(* PLC project EFBSH-649_PLC, ЗАО "Борисовский завод Металлист" CODESYS CODESYS V3.5 *)
(* stored: creationDateTime 2026-09-25T08:47:37, modificationDateTime 2026-09-25T08:47:37 *)

(* 8 регистров, адрес = 1100 + (индекс-1)*8 *)
TYPE ST_BunkerHmi :
STRUCT
    wSts      : WORD;   (* +0 маски GVL_Const.BS_* *)
    wAlm      : WORD;   (* +1 GVL_Const.BA_SF *)
    wBypass   : WORD;   (* +2 GVL_Const.BY_DVU *)
    uTDvu     : UINT;   (* +3 с *)
    uTRestart : UINT;   (* +4 с *)
    uRes5     : UINT;
    uRes6     : UINT;
    uRes7     : UINT;
END_STRUCT
END_TYPE

TYPE ST_BunkerIn :
STRUCT
    xDVU : BOOL;   (* 1 = верхний уровень *)
    xDNU : BOOL;   (* 1 = продукт на нижнем уровне (для бункера поз.27 - второй датчик) *)
    xSF  : BOOL;   (* станции TORBA: 1 = автомат пульта управления включен *)
END_STRUCT
END_TYPE

TYPE ST_BunkerPar :
STRUCT
    wBypass   : WORD;   (* GVL_Const.BY_DVU - ДВУ отключен *)
    uTDvu     : UINT;   (* задержка срабатывания ДВУ, с *)
    uTRestart : UINT;   (* задержка повторного пуска после снятия ДВУ, с *)
END_STRUCT
END_TYPE

(* Общий блок, %MW0..%MW31 *)
TYPE ST_GlobHmi :
STRUCT
    wCmd        : WORD;  (* +0  маски GVL_Const.G_* *)
    wSts        : WORD;  (* +1  маски GVL_Const.GS_* *)
    wAlm        : WORD;  (* +2  аварийные стопы 1..10 (биты 0..9), 10 пожар, 11 фазы *)
    wWarn       : WORD;  (* +3  маски GVL_Const.GW_* *)
    uHeartbeat  : UINT;  (* +4  счётчик секунд, контроль связи *)
    uTPreStart  : UINT;  (* +5  предпусковой сигнал, с *)
    uTDksGrace  : UINT;  (* +6  разгон до контроля ДКС, с *)
    uTDksPulse  : UINT;  (* +7  нет импульсов ДКС, 0.1 с *)
    uTFcFb      : UINT;  (* +8  нет сигнала работы ПЧ, с *)
    uTFsStart   : UINT;  (* +9  нет статуса фотосепаратора после пуска, с *)
    uTGateMove  : UINT;  (* +10 контроль хода заслонки поз.1, с *)
    uSirenOn    : UINT;  (* +11 1 = аварийная сирена разрешена *)
    uRes        : ARRAY[12..31] OF UINT;
END_STRUCT
END_TYPE

TYPE ST_GlobPar :
STRUCT
    uTPreStart : UINT;
    uTDksGrace : UINT;
    uTDksPulse : UINT;   (* 0.1 с *)
    uTFcFb     : UINT;
    uTFsStart  : UINT;
    uTGateMove : UINT;
    uSirenOn   : UINT;
END_STRUCT
END_TYPE

(* Связь "механизм подаёт на ..." для блокировок и последовательностей *)
TYPE ST_Link :
STRUCT
    iFrom    : INT;    (* индекс механизма-источника *)
    eTo      : INT;    (* GVL_Const.LT_MECH / LT_BUNKER / LT_INVALID *)
    iTo      : INT;    (* индекс механизма или бункера *)
    xProduct : BOOL;   (* TRUE - поток продукта (пауза по ДВУ распространяется назад),
                          FALSE - вспомогательная связь (аспирация, отходы) *)
END_STRUCT
END_TYPE

(* Постоянная конфигурация механизма *)
TYPE ST_MechCfg :
STRUCT
    eKind     : INT;     (* GVL_Const.K_DOL / K_FC / K_GATE / K_FS *)
    xHasQF    : BOOL;    (* контроль автомата защиты (QF/SF) *)
    eDks      : INT;     (* GVL_Const.DKS_NONE / DKS_PULSE / DKS_LEVEL *)
    xHasDSL   : BOOL;    (* датчики сбегания ленты 1 и 2 *)
    xHasDP    : BOOL;    (* датчик подпора *)
    xHasLocal : BOOL;    (* пост местного управления: ключ Авт/Ручн, Пуск, Стоп *)
    xHasEStop : BOOL;    (* аварийный/концевой стоп у механизма *)
    uDefTOn   : UINT;    (* задержка пуска по умолчанию, с *)
    uDefTOff  : UINT;    (* задержка останова по умолчанию, с *)
END_STRUCT
END_TYPE

(* Обмен с панелью по механизму: 16 регистров %MW (только 16-битные поля).
   Адрес = 200 + (индекс-1)*16 + смещение. *)
TYPE ST_MechHmi :
STRUCT
    wCmd           : WORD;  (* +0  команды панели, маски GVL_Const.C_* *)
    wSts           : WORD;  (* +1  состояние, маски GVL_Const.S_* *)
    wAlm           : WORD;  (* +2  аварии (с фиксацией), маски GVL_Const.A_* *)
    wBypass        : WORD;  (* +3  отключение датчиков (запись с паролем) *)
    uTOn           : UINT;  (* +4  задержка пуска, с *)
    uTOff          : UINT;  (* +5  задержка останова, с *)
    uToInterval    : UINT;  (* +6  интервал ТО, ч *)
    uHoursSinceTO  : UINT;  (* +7  наработка после ТО, ч *)
    uHoursTotal    : UINT;  (* +8  наработка всего, ч *)
    uMinutes       : UINT;  (* +9  минуты наработки (0..59) *)
    iState         : INT;   (* +10 0 стоп, 1 пуск, 2 работа, 3 останов, 4 авария, 5 местное *)
    uRes11         : UINT;
    uRes12         : UINT;
    uRes13         : UINT;
    uRes14         : UINT;
    uRes15         : UINT;
END_STRUCT
END_TYPE

(* Логические входы механизма (после учёта полярности в PRG_Inputs) *)
TYPE ST_MechIn :
STRUCT
    xQF       : BOOL;    (* 1 = автомат включен *)
    xDKS      : BOOL;    (* импульсы/уровень датчика контроля скорости *)
    xDSL1     : BOOL;    (* 1 = лента в норме *)
    xDSL2     : BOOL;
    xDP       : BOOL;    (* 1 = подпора нет *)
    xLocal    : BOOL;    (* 1 = ключ поста в положении "ручн." (местное управление) *)
    xLocStart : BOOL;    (* кнопка "Пуск" поста, НО *)
    xLocStop  : BOOL;    (* 1 = кнопка "Стоп" поста не нажата (НЗ) *)
    xEStop    : BOOL;    (* 1 = аварийный/концевой стоп не нажат (НЗ) *)
    xFcFault  : BOOL;    (* 1 = авария ПЧ *)
    xFcReady  : BOOL;    (* 1 = готовность/работа ПЧ *)
    xFb1      : BOOL;    (* заслонка: открыта;  фотосепаратор: статус "работа" *)
    xFb2      : BOOL;    (* заслонка: закрыта;  фотосепаратор: внешнее управление *)
    xErr      : BOOL;    (* фотосепаратор: критическая ошибка *)
    xLocOpen  : BOOL;    (* заслонка: кнопка "Открыть" поста *)
    xLocClose : BOOL;    (* заслонка: кнопка "Закрыть" поста *)
    xAux      : BOOL;    (* фотосепаратор: компрессор в работе (автомат включен) *)
END_STRUCT
END_TYPE

TYPE ST_MechOut :
STRUCT
    qRun    : BOOL;      (* пуск двигателя / пуск ПЧ *)
    qPower  : BOOL;      (* включить питание ПЧ (сетевой контактор) *)
    qReset  : BOOL;      (* сброс аварии ПЧ, импульс *)
    qOpen   : BOOL;      (* заслонка: открыть *)
    qClose  : BOOL;      (* заслонка: закрыть *)
    qOn     : BOOL;      (* фотосепаратор: импульс "Включить" *)
    qOff    : BOOL;      (* фотосепаратор: импульс "Выключить" *)
    qEnable : BOOL;      (* фотосепаратор: разрешить секции 1-3 *)
END_STRUCT
END_TYPE

(* Уставки и счётчики механизма, хранятся в RETAIN *)
TYPE ST_MechPar :
STRUCT
    uTOn         : UINT;     (* задержка пуска, с *)
    uTOff        : UINT;     (* задержка останова, с *)
    uToInterval  : UINT;     (* интервал ТО, ч; 0 = не контролировать *)
    wBypass      : WORD;     (* отключенные датчики, маски GVL_Const.BY_* *)
    udSecTotal   : UDINT;    (* наработка всего, с *)
    udSecSinceTO : UDINT;    (* наработка после ТО, с *)
END_STRUCT
END_TYPE

(* 4 регистра, адрес = 100 + (номер-1)*4 *)
TYPE ST_RouteHmi :
STRUCT
    wCmd      : WORD;  (* +0 маски GVL_Const.RC_* *)
    wSts      : WORD;  (* +1 маски GVL_Const.RS_* *)
    iNotReady : INT;   (* +2 причина отказа в пуске: 1..37 механизм, 101..105 клапан, 201..207 бункер,
                          -1 общая авария/цепь управления, -2 конфликт маршрутов, -3 ошибка конфигурации *)
    iState    : INT;   (* +3 0 стоп, 1 предпусковой сигнал, 2 перевод клапанов, 3 работа, 4 останов *)
END_STRUCT
END_TYPE

(* 8 регистров, адрес = 1000 + (индекс-1)*8 *)
TYPE ST_ValveHmi :
STRUCT
    wCmd   : WORD;   (* +0 маски GVL_Const.VC_* *)
    wSts   : WORD;   (* +1 маски GVL_Const.VS_* *)
    wAlm   : WORD;   (* +2 маски GVL_Const.VA_* *)
    uTMove : UINT;   (* +3 контроль времени перевода, с *)
    uRes4  : UINT;
    uRes5  : UINT;
    uRes6  : UINT;
    uRes7  : UINT;
END_STRUCT
END_TYPE

TYPE ST_ValveIn :
STRUCT
    xSF : BOOL;  (* 1 = автомат привода включен *)
    xS1 : BOOL;  (* датчик положения 1 *)
    xS2 : BOOL;  (* датчик положения 2 *)
END_STRUCT
END_TYPE

TYPE ST_ValveOut :
STRUCT
    q1 : BOOL;   (* перевод в положение 1 *)
    q2 : BOOL;   (* перевод в положение 2 *)
END_STRUCT
END_TYPE

TYPE ST_ValvePar :
STRUCT
    uTMove : UINT;   (* контроль времени перевода, с *)
END_STRUCT
END_TYPE

(* global variable list GVL *)
(* Рабочие переменные программы *)
VAR_GLOBAL
    (* ---- общие входы (заполняет PRG_Inputs) ---- *)
    xSysOnIn     : BOOL;                     (* 1K1: цепь управления включена *)
    aEStopIn     : ARRAY[1..10] OF BOOL;     (* 1 = аварийный стоп не нажат *)
    xFireOkIn    : BOOL;                     (* 1 = нет пожарной тревоги *)
    xPhaseOkIn   : BOOL;                     (* 1 = фазы в норме *)
    xFsAspPwrIn  : BOOL;
    xDryerOkIn   : BOOL;
    xComprOkIn   : BOOL;
    xCompr2OkIn  : BOOL;

    (* ---- общие флаги (PRG_System) ---- *)
    xSysOn     : BOOL;     (* цепь управления включена *)
    xGlobalOk  : BOOL;     (* цепь управления, аварийные стопы, пожар, фазы - в норме *)
    xReset     : BOOL;     (* импульс сброса аварий на один цикл *)
    xSetup     : BOOL;     (* режим наладки *)
    xStopAll   : BOOL;     (* импульс "остановить все маршруты" *)
    xPulse1s   : BOOL;     (* импульс раз в секунду на один цикл *)
    xBlink     : BOOL;     (* меандр 1 Гц *)
    xPreStart  : BOOL;     (* идёт предпусковой сигнал *)
    xAnyAlarm    : BOOL;
    xAnyNewAlarm : BOOL;
    qSiren     : BOOL;
    qLamp      : BOOL;

    (* ---- механизмы ---- *)
    aMechIn   : ARRAY[1..GVL_Const.N_MECH] OF ST_MechIn;
    aMechOut  : ARRAY[1..GVL_Const.N_MECH] OF ST_MechOut;
    aRun      : ARRAY[1..GVL_Const.N_MECH] OF BOOL;   (* механизм работает *)
    aReady    : ARRAY[1..GVL_Const.N_MECH] OF BOOL;   (* готов к работе в маршруте *)
    aAuto     : ARRAY[1..GVL_Const.N_MECH] OF BOOL;   (* в автоматическом режиме *)
    aAlarm    : ARRAY[1..GVL_Const.N_MECH] OF BOOL;
    aDemand   : ARRAY[1..GVL_Const.N_MECH] OF BOOL;   (* требуется активным маршрутом *)
    aPredRun  : ARRAY[1..GVL_Const.N_MECH] OF BOOL;   (* работает механизм, подающий на данный *)
    aSuccAuto : ARRAY[1..GVL_Const.N_MECH] OF BOOL;   (* все последующие механизмы работают *)
    aSuccMan  : ARRAY[1..GVL_Const.N_MECH] OF BOOL;   (* то же + бункеры на выходе не полны *)
    aBlocked  : ARRAY[1..GVL_Const.N_MECH] OF BOOL;   (* участок стоит на паузе по ДВУ *)

    (* ---- переключатели потока ---- *)
    aValveIn     : ARRAY[1..GVL_Const.N_VALVE] OF ST_ValveIn;
    aValveOut    : ARRAY[1..GVL_Const.N_VALVE] OF ST_ValveOut;
    aValvePos    : ARRAY[1..GVL_Const.N_VALVE] OF INT;   (* 0 - не определено, 1, 2 *)
    aValveTarget : ARRAY[1..GVL_Const.N_VALVE] OF INT;   (* задание от маршрутов *)
    aValveReady  : ARRAY[1..GVL_Const.N_VALVE] OF BOOL;
    aValveAlarm  : ARRAY[1..GVL_Const.N_VALVE] OF BOOL;

    (* ---- бункеры ---- *)
    aBunkerIn    : ARRAY[1..GVL_Const.N_BUNKER] OF ST_BunkerIn;
    aBunkerFull  : ARRAY[1..GVL_Const.N_BUNKER] OF BOOL;
    aBunkerAlarm : ARRAY[1..GVL_Const.N_BUNKER] OF BOOL;

    (* ---- связи и маршруты ---- *)
    aLinks       : ARRAY[1..GVL_Const.N_LINK] OF ST_Link;
    nLinks       : INT;
    aMember      : ARRAY[1..GVL_Const.N_ROUTE, 1..GVL_Const.N_MECH] OF BOOL;    (* состав маршрута *)
    aMemberB     : ARRAY[1..GVL_Const.N_ROUTE, 1..GVL_Const.N_BUNKER] OF BOOL;  (* бункеры маршрута *)
    aRouteCfgErr : ARRAY[1..GVL_Const.N_ROUTE] OF BOOL;
    aRouteState  : ARRAY[1..GVL_Const.N_ROUTE] OF INT;
    aRouteFault  : ARRAY[1..GVL_Const.N_ROUTE] OF BOOL;
END_VAR

(* global variable list GVL_Const *)
(* Константы проекта ЕФБШ-649.01-АТХ, ЛПЗС-5 ССЦ "Золотой початок".
   Номера позиций "поз." - по технологической схеме (Приложение 1). *)
VAR_GLOBAL CONSTANT
    N_MECH   : INT := 37;
    N_VALVE  : INT := 5;
    N_BUNKER : INT := 7;
    N_ROUTE  : INT := 11;
    N_LINK   : INT := 64;
    N_HEAD   : INT := 6;

    (* ---- механизмы (индекс = номер в панели) ---- *)
    M_GATE1    : INT := 1;   (* заслонка бункера растаривания поз.1, ПЧ 51UZ1 *)
    M_N3       : INT := 2;   (* нория поз.3 *)
    M_MUZ5_FD  : INT := 3;   (* МУЗ-8М поз.5 - битер (питатель), ПЧ 5UZ1 *)
    M_MUZ5     : INT := 4;   (* МУЗ-8М поз.5 - основной двигатель *)
    M_FAN6     : INT := 5;   (* вентилятор аспирации поз.6 *)
    M_SL6      : INT := 6;   (* шлюзовой затвор поз.6 *)
    M_N7       : INT := 7;   (* нория поз.7 *)
    M_TOR9_FD  : INT := 8;   (* ТОР-18 поз.9 - двигатель 0,75 кВт, ПЧ 11UZ1 *)
    M_TOR9     : INT := 9;   (* ТОР-18 поз.9 - основной двигатель *)
    M_FAN10    : INT := 10;  (* вентилятор аспирации поз.10 *)
    M_SL10     : INT := 11;  (* шлюзовой затвор поз.10 *)
    M_N11      : INT := 12;  (* нория поз.11 *)
    M_BT14_1   : INT := 13;  (* блок триерный БТ-9/2 поз.14 - двигатель 1, ПЧ 24UZ1 *)
    M_BT14_2   : INT := 14;  (* блок триерный БТ-9/2 поз.14 - двигатель 2, ПЧ 25UZ1 *)
    M_N16      : INT := 15;  (* нория поз.16 *)
    M_KSP18_FD : INT := 16;  (* КСП-11М поз.18 - битер (питатель), ПЧ 29UZ1 *)
    M_KSP18    : INT := 17;  (* КСП-11М поз.18 - основной двигатель *)
    M_FAN19    : INT := 18;  (* вентилятор аспирации поз.19 *)
    M_SL19     : INT := 19;  (* шлюзовой затвор поз.19 *)
    M_N20      : INT := 20;  (* нория поз.20 *)
    M_N21      : INT := 21;  (* нория поз.21 *)
    M_SP24_DRV : INT := 22;  (* СП-200 поз.24 - привод деки, ПЧ 36UZ1 *)
    M_SP24_FAN : INT := 23;  (* СП-200 поз.24 - вентилятор стола 11 кВт (звезда-треугольник) *)
    M_FAN25    : INT := 24;  (* вентилятор аспирации поз.25 *)
    M_SL25     : INT := 25;  (* шлюзовой затвор поз.25 *)
    M_ZN26     : INT := 26;  (* Z-нория поз.26, ПЧ 48UZ1 *)
    M_FS27     : INT := 27;  (* фотосепаратор СмартСорт поз.27 *)
    M_FAN28    : INT := 28;  (* вентилятор аспирации поз.28 *)
    M_SL28     : INT := 29;  (* шлюзовой затвор поз.28 *)
    M_ZN29     : INT := 30;  (* Z-нория поз.29, ПЧ 50UZ1 *)
    M_SH30     : INT := 31;  (* конвейер шнековый КШ-4-150 поз.30 *)
    M_SH31     : INT := 32;  (* конвейер шнековый КШU-150 поз.31 *)
    M_SH32     : INT := 33;  (* конвейер шнековый КШU-150 поз.32 *)
    M_SH33     : INT := 34;  (* конвейер шнековый КШU-150 поз.33 *)
    M_KC34     : INT := 35;  (* конвейер цепной КЦСВ поз.34 *)
    M_KC35     : INT := 36;  (* конвейер цепной КЦСН поз.35 *)
    M_KC36     : INT := 37;  (* конвейер цепной КЦСН поз.36 *)

    (* ---- переключатели потока (положение 1 / положение 2) ---- *)
    V_V12_1 : INT := 1;   (* поз.12(1): 1 - на TORBA поз.13(1),  2 - на поз.12(2) *)
    V_V12_2 : INT := 2;   (* поз.12(2): 1 - на БТ поз.14,         2 - на растариватель 15(1) -> нория 16 *)
    V_V12_3 : INT := 3;   (* поз.12(3): 1 - на бункер поз.17 (КСП), 2 - на норию поз.20 *)
    V_V12_4 : INT := 4;   (* поз.12(4): 1 - на бункер поз.22 (СП),  2 - на Z-норию поз.26 *)
    V_V49   : INT := 5;   (* выгрузка Z-нории поз.26: 1 - включена (на TORBA 13(2)), 2 - выключена (на ФС поз.27) *)

    (* ---- бункеры ---- *)
    B_B4    : INT := 1;   (* бункер оперативный поз.4 *)
    B_B8    : INT := 2;   (* бункер оперативный поз.8 *)
    B_B17   : INT := 3;   (* бункер оперативный поз.17 *)
    B_B22   : INT := 4;   (* бункер оперативный поз.22 *)
    B_B27   : INT := 5;   (* приёмный бункер фотосепаратора поз.27 *)
    B_T13_1 : INT := 6;   (* станция затаривания TORBA-1000 поз.13(1) *)
    B_T13_2 : INT := 7;   (* станция затаривания TORBA-1000 поз.13(2) *)

    (* ---- типы механизмов ---- *)
    K_DOL  : INT := 0;    (* прямой пуск *)
    K_FC   : INT := 1;    (* частотный преобразователь: питание, пуск, сброс *)
    K_GATE : INT := 2;    (* заслонка с ПЧ: открыть/закрыть, концевики *)
    K_FS   : INT := 3;    (* фотосепаратор: импульсы вкл/выкл, разрешение секций *)

    DKS_NONE  : INT := 0;
    DKS_PULSE : INT := 1; (* индуктивный датчик, импульсы *)
    DKS_LEVEL : INT := 2; (* реле движения РДД-03, уровень 1 = движение есть *)

    MODE_AUTO  : INT := 0;
    MODE_MAN   : INT := 1;
    MODE_LOCAL : INT := 2;

    LT_MECH    : INT := 0;
    LT_BUNKER  : INT := 1;
    LT_INVALID : INT := 2; (* клапан не в положении - подача не определена *)

    RST_IDLE     : INT := 0;
    RST_PRESTART : INT := 1;
    RST_VALVES   : INT := 2;
    RST_RUN      : INT := 3;
    RST_STOPPING : INT := 4;

    (* ---- полярность датчиков (проверить при ПНР) ---- *)
    CFG_DSL_OK      : BOOL := TRUE;   (* ДСЛ И25-NO/NC: 1 = лента в норме *)
    CFG_DP_OK       : BOOL := TRUE;   (* ДП норий Е13-NC: 1 = подпора нет *)
    CFG_DP_SCREW_OK : BOOL := TRUE;   (* ДП шнеков, концевик EMAS: 1 = подпора нет *)
    CFG_DP_CHAIN_OK : BOOL := FALSE;  (* ДП цепных конвейеров через реле РСУ-4 (KM3 13-14): 1 = подпор *)
    CFG_DVU_FULL    : BOOL := TRUE;   (* ДВУ через промежуточное реле: 1 = бункер полон *)
    CFG_DNU_ON      : BOOL := TRUE;   (* ДНУ: 1 = продукт есть *)
    CFG_FC_FAULT    : BOOL := TRUE;   (* реле аварии ПЧ Hope530 (1TA-1TC): 1 = авария *)
    CFG_SA_LOCAL    : BOOL := TRUE;   (* ключ поста "Автом./ручн." (11-14): 1 = ручн. (местное) *)

    (* ---- команды механизма (ST_MechHmi.wCmd) ---- *)
    C_START    : WORD := 16#0001;   (* пуск в ручном режиме, импульс *)
    C_STOP     : WORD := 16#0002;   (* стоп в ручном режиме, импульс *)
    C_MANUAL   : WORD := 16#0004;   (* 1 = ручной режим с панели, 0 = автомат *)
    C_RESET_TO : WORD := 16#0008;   (* сброс счётчика ТО, импульс *)
    C_OPEN     : WORD := 16#0010;   (* заслонка: открывать, пока нажато *)
    C_CLOSE    : WORD := 16#0020;   (* заслонка: закрывать, пока нажато *)

    (* ---- состояние механизма (ST_MechHmi.wSts) ---- *)
    S_RUN      : WORD := 16#0001;
    S_CMD      : WORD := 16#0002;
    S_READY    : WORD := 16#0004;
    S_ALARM    : WORD := 16#0008;
    S_LOCAL    : WORD := 16#0010;
    S_MANUAL   : WORD := 16#0020;
    S_SETUP    : WORD := 16#0040;
    S_STARTING : WORD := 16#0080;
    S_STOPPING : WORD := 16#0100;
    S_DEMAND   : WORD := 16#0200;
    S_PAUSE    : WORD := 16#0400;
    S_TO_DUE   : WORD := 16#0800;
    S_OPENED   : WORD := 16#1000;
    S_CLOSED   : WORD := 16#2000;
    S_SEQ_TRIP : WORD := 16#4000;   (* остановлен блокировкой: встал последующий механизм *)
    S_SUCC_OK  : WORD := 16#8000;   (* последующие механизмы в работе - ручной пуск разрешён *)

    (* ---- аварии механизма (ST_MechHmi.wAlm) ---- *)
    A_QF      : WORD := 16#0001;    (* защита двигателя / ПЧ *)
    A_DKS     : WORD := 16#0002;    (* нет вращения (ДКС) *)
    A_DSL1    : WORD := 16#0004;    (* сбег ленты 1 *)
    A_DSL2    : WORD := 16#0008;    (* сбег ленты 2 *)
    A_DP      : WORD := 16#0010;    (* подпор *)
    A_ESTOP   : WORD := 16#0020;    (* аварийный / концевой стоп у механизма *)
    A_LOCSTOP : WORD := 16#0040;    (* нажат местный "Стоп" при работе от панели *)
    A_FC      : WORD := 16#0080;    (* авария ПЧ *)
    A_FCFB    : WORD := 16#0100;    (* нет сигнала работы ПЧ *)
    A_MOVE    : WORD := 16#0200;    (* заслонка не дошла за заданное время *)
    A_POS     : WORD := 16#0400;    (* заслонка: оба концевика *)
    A_FSERR   : WORD := 16#0800;    (* фотосепаратор: критическая ошибка *)
    A_FSFB    : WORD := 16#1000;    (* фотосепаратор: нет статуса работы *)
    A_HARD    : WORD := 16#08A1;    (* аварии, которые не отключаются в режиме наладки: QF, ESTOP, FC, FSERR *)

    (* ---- отключение датчиков (ST_MechHmi.wBypass / ST_BunkerHmi.wBypass) ---- *)
    BY_DKS  : WORD := 16#0001;
    BY_DSL1 : WORD := 16#0002;
    BY_DSL2 : WORD := 16#0004;
    BY_DP   : WORD := 16#0008;
    BY_AUX  : WORD := 16#0010;      (* фотосепаратор: не требовать работу компрессора *)
    BY_DVU  : WORD := 16#0001;      (* бункер: ДВУ отключен *)

    (* ---- переключатели потока ---- *)
    VC_POS1   : WORD := 16#0001;    (* перевести в положение 1, импульс (ручной режим) *)
    VC_POS2   : WORD := 16#0002;
    VC_MANUAL : WORD := 16#0004;
    VS_POS1   : WORD := 16#0001;
    VS_POS2   : WORD := 16#0002;
    VS_MOVING : WORD := 16#0004;
    VS_ALARM  : WORD := 16#0008;
    VS_MANUAL : WORD := 16#0010;
    VS_ROUTE  : WORD := 16#0020;    (* положение задано маршрутом *)
    VS_FLOW   : WORD := 16#0040;    (* подающий механизм работает - ручной перевод запрещён *)
    VA_SF      : WORD := 16#0001;
    VA_TIMEOUT : WORD := 16#0002;
    VA_BOTH    : WORD := 16#0004;

    (* ---- бункеры ---- *)
    BS_DVU    : WORD := 16#0001;    (* ДВУ сработал (без задержки) *)
    BS_FULL   : WORD := 16#0002;    (* бункер полон - пауза подачи *)
    BS_DNU    : WORD := 16#0004;
    BS_BYPASS : WORD := 16#0008;
    BS_ALARM  : WORD := 16#0010;
    BA_SF     : WORD := 16#0001;    (* TORBA: отключен автомат пульта управления *)

    (* ---- маршруты ---- *)
    RC_TOGGLE : WORD := 16#0001;    (* "ПУСК" / повторное нажатие - "СТОП" *)
    RC_STOP   : WORD := 16#0002;
    RS_ACTIVE   : WORD := 16#0001;
    RS_PRESTART : WORD := 16#0002;
    RS_VALVES   : WORD := 16#0004;
    RS_RUN      : WORD := 16#0008;
    RS_STOPPING : WORD := 16#0010;
    RS_PAUSED   : WORD := 16#0020;
    RS_FAULT    : WORD := 16#0040;
    RS_NOTREADY : WORD := 16#0080;
    RS_CONFLICT : WORD := 16#0100;
    RS_ALLRUN   : WORD := 16#0200;

    (* ---- общий блок ---- *)
    G_RESET   : WORD := 16#0001;    (* сброс аварий, импульс (после подтверждения на панели) *)
    G_MUTE    : WORD := 16#0002;    (* отключить звук сирены, импульс *)
    G_SETUP   : WORD := 16#0004;    (* режим наладки (панель выставляет после ввода пароля) *)
    G_STOPALL : WORD := 16#0008;    (* остановить все маршруты, импульс *)
    GS_SYSON    : WORD := 16#0001;  (* цепь управления включена (1K1) *)
    GS_OK       : WORD := 16#0002;  (* нет общих аварий *)
    GS_ALARM    : WORD := 16#0004;  (* есть активные аварии *)
    GS_SIREN    : WORD := 16#0008;
    GS_SETUP    : WORD := 16#0010;
    GS_PRESTART : WORD := 16#0020;
    GA_FIRE  : WORD := 16#0400;
    GA_PHASE : WORD := 16#0800;
    GW_COMPR  : WORD := 16#0001;    (* отключен автомат компрессора 57SF1 *)
    GW_COMPR2 : WORD := 16#0002;    (* 58QF1 (опция) *)
    GW_DRYER  : WORD := 16#0004;    (* 56SF1 (опция) *)
    GW_FSASP  : WORD := 16#0008;    (* 53SF1 питание аспирации ФС (опция) *)
    GW_SYSOFF : WORD := 16#0010;    (* цепь управления отключена *)

    T_MAX_S  : UINT := 3600;
    RETAIN_MAGIC : UINT := 16#6491;

    (* ---- конфигурация механизмов ---- *)
    MECH_CFG : ARRAY[1..37] OF ST_MechCfg := [
        (eKind := 2, xHasQF := TRUE, eDks := 0, xHasDSL := FALSE, xHasDP := FALSE, xHasLocal := TRUE,  xHasEStop := FALSE, uDefTOn := 2,  uDefTOff := 0),   (* 1  заслонка поз.1 *)
        (eKind := 0, xHasQF := TRUE, eDks := 1, xHasDSL := TRUE,  xHasDP := TRUE,  xHasLocal := TRUE,  xHasEStop := TRUE,  uDefTOn := 3,  uDefTOff := 10),  (* 2  нория поз.3 *)
        (eKind := 1, xHasQF := TRUE, eDks := 0, xHasDSL := FALSE, xHasDP := FALSE, xHasLocal := FALSE, xHasEStop := TRUE,  uDefTOn := 3,  uDefTOff := 0),   (* 3  битер МУЗ *)
        (eKind := 0, xHasQF := TRUE, eDks := 0, xHasDSL := FALSE, xHasDP := FALSE, xHasLocal := FALSE, xHasEStop := FALSE, uDefTOn := 5,  uDefTOff := 15),  (* 4  МУЗ-8М *)
        (eKind := 0, xHasQF := TRUE, eDks := 0, xHasDSL := FALSE, xHasDP := FALSE, xHasLocal := FALSE, xHasEStop := FALSE, uDefTOn := 5,  uDefTOff := 30),  (* 5  вентилятор поз.6 *)
        (eKind := 0, xHasQF := TRUE, eDks := 1, xHasDSL := FALSE, xHasDP := FALSE, xHasLocal := FALSE, xHasEStop := FALSE, uDefTOn := 3,  uDefTOff := 40),  (* 6  шлюз поз.6 *)
        (eKind := 0, xHasQF := TRUE, eDks := 1, xHasDSL := TRUE,  xHasDP := TRUE,  xHasLocal := TRUE,  xHasEStop := TRUE,  uDefTOn := 3,  uDefTOff := 10),  (* 7  нория поз.7 *)
        (eKind := 1, xHasQF := TRUE, eDks := 0, xHasDSL := FALSE, xHasDP := FALSE, xHasLocal := FALSE, xHasEStop := TRUE,  uDefTOn := 3,  uDefTOff := 0),   (* 8  ПЧ ТОР-18 *)
        (eKind := 0, xHasQF := TRUE, eDks := 0, xHasDSL := FALSE, xHasDP := FALSE, xHasLocal := FALSE, xHasEStop := FALSE, uDefTOn := 5,  uDefTOff := 15),  (* 9  ТОР-18 *)
        (eKind := 0, xHasQF := TRUE, eDks := 0, xHasDSL := FALSE, xHasDP := FALSE, xHasLocal := FALSE, xHasEStop := FALSE, uDefTOn := 5,  uDefTOff := 30),  (* 10 вентилятор поз.10 *)
        (eKind := 0, xHasQF := TRUE, eDks := 1, xHasDSL := FALSE, xHasDP := FALSE, xHasLocal := FALSE, xHasEStop := FALSE, uDefTOn := 3,  uDefTOff := 40),  (* 11 шлюз поз.10 *)
        (eKind := 0, xHasQF := TRUE, eDks := 1, xHasDSL := TRUE,  xHasDP := TRUE,  xHasLocal := TRUE,  xHasEStop := TRUE,  uDefTOn := 3,  uDefTOff := 10),  (* 12 нория поз.11 *)
        (eKind := 1, xHasQF := TRUE, eDks := 0, xHasDSL := FALSE, xHasDP := FALSE, xHasLocal := FALSE, xHasEStop := TRUE,  uDefTOn := 5,  uDefTOff := 15),  (* 13 БТ-9/2 двигатель 1 *)
        (eKind := 1, xHasQF := TRUE, eDks := 0, xHasDSL := FALSE, xHasDP := FALSE, xHasLocal := FALSE, xHasEStop := TRUE,  uDefTOn := 5,  uDefTOff := 15),  (* 14 БТ-9/2 двигатель 2 *)
        (eKind := 0, xHasQF := TRUE, eDks := 1, xHasDSL := TRUE,  xHasDP := TRUE,  xHasLocal := TRUE,  xHasEStop := TRUE,  uDefTOn := 3,  uDefTOff := 10),  (* 15 нория поз.16 *)
        (eKind := 1, xHasQF := TRUE, eDks := 0, xHasDSL := FALSE, xHasDP := FALSE, xHasLocal := FALSE, xHasEStop := TRUE,  uDefTOn := 3,  uDefTOff := 0),   (* 16 битер КСП *)
        (eKind := 0, xHasQF := TRUE, eDks := 0, xHasDSL := FALSE, xHasDP := FALSE, xHasLocal := FALSE, xHasEStop := FALSE, uDefTOn := 5,  uDefTOff := 15),  (* 17 КСП-11М *)
        (eKind := 0, xHasQF := TRUE, eDks := 0, xHasDSL := FALSE, xHasDP := FALSE, xHasLocal := FALSE, xHasEStop := FALSE, uDefTOn := 5,  uDefTOff := 30),  (* 18 вентилятор поз.19 *)
        (eKind := 0, xHasQF := TRUE, eDks := 1, xHasDSL := FALSE, xHasDP := FALSE, xHasLocal := FALSE, xHasEStop := FALSE, uDefTOn := 3,  uDefTOff := 40),  (* 19 шлюз поз.19 *)
        (eKind := 0, xHasQF := TRUE, eDks := 1, xHasDSL := TRUE,  xHasDP := TRUE,  xHasLocal := TRUE,  xHasEStop := TRUE,  uDefTOn := 3,  uDefTOff := 10),  (* 20 нория поз.20 *)
        (eKind := 0, xHasQF := TRUE, eDks := 1, xHasDSL := TRUE,  xHasDP := TRUE,  xHasLocal := TRUE,  xHasEStop := TRUE,  uDefTOn := 3,  uDefTOff := 10),  (* 21 нория поз.21 *)
        (eKind := 1, xHasQF := TRUE, eDks := 0, xHasDSL := FALSE, xHasDP := FALSE, xHasLocal := FALSE, xHasEStop := TRUE,  uDefTOn := 5,  uDefTOff := 10),  (* 22 СП-200 привод *)
        (eKind := 0, xHasQF := TRUE, eDks := 0, xHasDSL := FALSE, xHasDP := FALSE, xHasLocal := FALSE, xHasEStop := FALSE, uDefTOn := 10, uDefTOff := 15),  (* 23 СП-200 вентилятор *)
        (eKind := 0, xHasQF := TRUE, eDks := 0, xHasDSL := FALSE, xHasDP := FALSE, xHasLocal := FALSE, xHasEStop := FALSE, uDefTOn := 5,  uDefTOff := 30),  (* 24 вентилятор поз.25 *)
        (eKind := 0, xHasQF := TRUE, eDks := 1, xHasDSL := FALSE, xHasDP := FALSE, xHasLocal := FALSE, xHasEStop := FALSE, uDefTOn := 3,  uDefTOff := 40),  (* 25 шлюз поз.25 *)
        (eKind := 1, xHasQF := TRUE, eDks := 1, xHasDSL := FALSE, xHasDP := FALSE, xHasLocal := TRUE,  xHasEStop := TRUE,  uDefTOn := 3,  uDefTOff := 10),  (* 26 Z-нория поз.26 *)
        (eKind := 3, xHasQF := TRUE, eDks := 0, xHasDSL := FALSE, xHasDP := FALSE, xHasLocal := FALSE, xHasEStop := FALSE, uDefTOn := 5,  uDefTOff := 10),  (* 27 фотосепаратор *)
        (eKind := 0, xHasQF := TRUE, eDks := 0, xHasDSL := FALSE, xHasDP := FALSE, xHasLocal := FALSE, xHasEStop := FALSE, uDefTOn := 5,  uDefTOff := 30),  (* 28 вентилятор поз.28 *)
        (eKind := 0, xHasQF := TRUE, eDks := 1, xHasDSL := FALSE, xHasDP := FALSE, xHasLocal := FALSE, xHasEStop := FALSE, uDefTOn := 3,  uDefTOff := 40),  (* 29 шлюз поз.28 *)
        (eKind := 1, xHasQF := TRUE, eDks := 1, xHasDSL := FALSE, xHasDP := FALSE, xHasLocal := TRUE,  xHasEStop := TRUE,  uDefTOn := 3,  uDefTOff := 10),  (* 30 Z-нория поз.29 *)
        (eKind := 0, xHasQF := TRUE, eDks := 0, xHasDSL := FALSE, xHasDP := FALSE, xHasLocal := TRUE,  xHasEStop := TRUE,  uDefTOn := 3,  uDefTOff := 30),  (* 31 шнек поз.30 (ДКС, ДП - опция) *)
        (eKind := 0, xHasQF := TRUE, eDks := 1, xHasDSL := FALSE, xHasDP := TRUE,  xHasLocal := TRUE,  xHasEStop := TRUE,  uDefTOn := 3,  uDefTOff := 30),  (* 32 шнек поз.31 *)
        (eKind := 0, xHasQF := TRUE, eDks := 1, xHasDSL := FALSE, xHasDP := TRUE,  xHasLocal := TRUE,  xHasEStop := TRUE,  uDefTOn := 3,  uDefTOff := 30),  (* 33 шнек поз.32 *)
        (eKind := 0, xHasQF := TRUE, eDks := 1, xHasDSL := FALSE, xHasDP := TRUE,  xHasLocal := TRUE,  xHasEStop := TRUE,  uDefTOn := 3,  uDefTOff := 30),  (* 34 шнек поз.33 *)
        (eKind := 0, xHasQF := TRUE, eDks := 2, xHasDSL := FALSE, xHasDP := TRUE,  xHasLocal := TRUE,  xHasEStop := TRUE,  uDefTOn := 3,  uDefTOff := 30),  (* 35 цепной поз.34 *)
        (eKind := 0, xHasQF := TRUE, eDks := 2, xHasDSL := FALSE, xHasDP := TRUE,  xHasLocal := TRUE,  xHasEStop := TRUE,  uDefTOn := 3,  uDefTOff := 30),  (* 36 цепной поз.35 *)
        (eKind := 0, xHasQF := TRUE, eDks := 2, xHasDSL := FALSE, xHasDP := TRUE,  xHasLocal := TRUE,  xHasEStop := TRUE,  uDefTOn := 3,  uDefTOff := 30)   (* 37 цепной поз.36 *)
    ];

    (* ---- маршруты (Приложение 5) ----
       1  Очистка: воронка - ... - БТ - нория 16 - нория 20 - СП - Z26 - ФС - Z29 - TORBA 13(2) (мимо КСП)
       2  Очистка мимо БТ (через КСП)
       3  Очистка мимо БТ и КСП
       4  Очистка мимо КСП и фотосепаратора
       5  Очистка мимо БТ, КСП и фотосепаратора
       6  Воронка - ... - ТОР - нория 11 - TORBA 13(1)
       7  Растариватель 15(1) - нория 16 - КСП - нория 20 - СП - Z26 - ФС - Z29 - TORBA 13(2)
       8  Растариватель 15(1) - нория 16 - КСП - нория 20 - СП - Z26 - TORBA 13(2)
       9  Растариватель 15(2) - нория 21 - СП - Z26 - ФС - Z29 - TORBA 13(2)
       10 Растариватель 15(2) - нория 21 - СП - Z26 - TORBA 13(2)
       11 Растариватель 15(2) - нория 21 - Z26 - ФС - Z29 - TORBA 13(2)
       Головные механизмы участков (от которых по связям определяется состав маршрута):
       1 заслонка, 3 битер МУЗ, 8 ПЧ ТОР, 15 нория 16, 16 битер КСП, 21 нория 21, 22 привод СП, 27 ФС *)
    ROUTE_HEAD : ARRAY[1..11, 1..6] OF INT := [
        1, 3, 8, 22, 27, 0,
        1, 3, 8, 16, 22, 27,
        1, 3, 8, 22, 27, 0,
        1, 3, 8, 22, 0, 0,
        1, 3, 8, 22, 0, 0,
        1, 3, 8, 0, 0, 0,
        15, 16, 22, 27, 0, 0,
        15, 16, 22, 0, 0, 0,
        21, 22, 27, 0, 0, 0,
        21, 22, 0, 0, 0, 0,
        21, 27, 0, 0, 0, 0
    ];
    (* положения клапанов: 12(1), 12(2), 12(3), 12(4), выгрузка Z26; 0 = не участвует *)
    ROUTE_VALVE : ARRAY[1..11, 1..5] OF INT := [
        2, 1, 2, 0, 2,
        2, 2, 1, 0, 2,
        2, 2, 2, 0, 2,
        2, 1, 2, 0, 1,
        2, 2, 2, 0, 1,
        1, 0, 0, 0, 0,
        0, 0, 1, 0, 2,
        0, 0, 1, 0, 1,
        0, 0, 0, 1, 2,
        0, 0, 0, 1, 1,
        0, 0, 0, 2, 2
    ];
    (* запреты одновременного пуска (Приложение 5), TRUE = запрет *)
    ROUTE_CONFLICT : ARRAY[1..11, 1..11] OF BOOL := [
        55(TRUE),
        5(TRUE), 6(FALSE),
        5(TRUE), FALSE, 5(TRUE),
        5(TRUE), FALSE, 5(TRUE),
        5(TRUE), FALSE, 5(TRUE),
        5(TRUE), FALSE, 5(TRUE),
        5(TRUE), FALSE, 5(TRUE)
    ];

    (* механизм, подающий продукт на клапан (при его работе ручной перевод запрещён) *)
    VALVE_FEEDER : ARRAY[1..5] OF INT := [12, 12, 15, 21, 26];
    VALVE_HAS_SF : ARRAY[1..5] OF BOOL := [TRUE, TRUE, TRUE, TRUE, FALSE];
    BUNKER_HAS_SF : ARRAY[1..7] OF BOOL := [FALSE, FALSE, FALSE, FALSE, FALSE, TRUE, TRUE];
END_VAR

(* global variable list GVL_HMI *)
(* Обмен с панелью Weintek cMT2166X по Modbus TCP (регистры хранения = %MW контроллера).
   Карта регистров - doc/HMI_map.md. *)
VAR_GLOBAL
    stHmiG     AT %MW0    : ST_GlobHmi;                                    (* %MW0..31 *)
    aHmiRoute  AT %MW100  : ARRAY[1..GVL_Const.N_ROUTE] OF ST_RouteHmi;    (* %MW100..143, по 4 *)
    aHmiMech   AT %MW200  : ARRAY[1..GVL_Const.N_MECH] OF ST_MechHmi;      (* %MW200..791, по 16 *)
    aHmiValve  AT %MW1000 : ARRAY[1..GVL_Const.N_VALVE] OF ST_ValveHmi;    (* %MW1000..1039, по 8 *)
    aHmiBunker AT %MW1100 : ARRAY[1..GVL_Const.N_BUNKER] OF ST_BunkerHmi;  (* %MW1100..1155, по 8 *)
END_VAR

(* global variable list GVL_IO *)
(* Сгенерировано gen/gen_io.py из Э3 ЕФБШ-649.01-АТХ. Не редактировать вручную.
   Привязка к каналам: Machine Expert -> модуль -> "Соотнесение входов/выходов" (I/O Mapping) ->
   переменная канала = Application.GVL_IO.<имя> (см. doc/IO_map.csv). *)
VAR_GLOBAL
    (* ---- A1 TM241CE40T ---- *)
    DI_SYS_ON           : BOOL; (* A1 I0 [X0] Пуск системы; 1K1 (31-34); Шкаф управления — общие сигналы; лист 3 *)
    DI_ESTOP_1          : BOOL; (* A1 I1 [X1] Аварийный стоп (шкаф); 1K2 (21-24); Шкаф управления — общие сигналы; лист 3 *)
    DI_ESTOP_2          : BOOL; (* A1 I2 [X2] Аварийный стоп цех; 1K3 (21-24); Шкаф управления — общие сигналы; лист 3 *)
    DI_ESTOP_3          : BOOL; (* A1 I3 [X3] Аварийный стоп у МУЗ-8М (поз. 5); 1K4 (21-24); Шкаф управления — общие сигналы; лист 3 *)
    DI_ESTOP_4          : BOOL; (* A1 I4 [X4] Аварийный стоп у ТОР-18 (поз. 9); 1K5 (21-24); Шкаф управления — общие сигналы; лист 3 *)
    DI_ESTOP_5          : BOOL; (* A1 I5 [X5] Аварийный стоп у СП-200 (поз. 24); 1K6 (21-24); Шкаф управления — общие сигналы; лист 3 *)
    DI_ESTOP_6          : BOOL; (* A1 I6 [X6] Аварийный стоп у аспирации; 1K7 (21-24); Шкаф управления — общие сигналы; лист 3 *)
    DI_ESTOP_7          : BOOL; (* A1 I7 [X7] Аварийный стоп у фотосепаратора (поз. 27); 1K8 (21-24); Шкаф управления — общие сигналы; лист 3 *)
    DI_ESTOP_8          : BOOL; (* A1 I8 [X8] Аварийный стоп цех; 1K9 (21-24); Шкаф управления — общие сигналы; лист 3 *)
    DI_ESTOP_9          : BOOL; (* A1 I9 [X9] Аварийный стоп у выгрузки (поз. 13); 1K10 (21-24); Шкаф управления — общие сигналы; лист 3 *)
    DI_ESTOP_10         : BOOL; (* A1 I10 [X10] Аварийный стоп у нории верх (поз. 26); 1K11 (21-24); Шкаф управления — общие сигналы; лист 3 *)
    DI_FIRE_OK          : BOOL; (* A1 I11 [X11] Пожарная сигнализация; 1K12 (21-24); Шкаф управления — общие сигналы; лист 3 *)
    DI_PHASE_OK         : BOOL; (* A1 I12 [X12] Контроль фаз; 1KV1 (клемма 18); Шкаф управления — общие сигналы; лист 3 *)
    DI_A1_I13_RES       : BOOL; (* A1 I13 [X13] Резерв; 1K13 (21-24); Шкаф управления — общие сигналы; лист 3 *)
    DI_N3_DKS           : BOOL; (* A1 I14 [X14] ДКС; 2SR1; Нория НС-А.20.09 (поз. 3); лист 4 *)
    DI_N3_DSL1          : BOOL; (* A1 I15 [X15] Датчик сбега ленты 1; 2SQ1; Нория НС-А.20.09 (поз. 3); лист 4 *)
    DI_N3_DSL2          : BOOL; (* A1 I16 [X16] Датчик сбега ленты 2; 2SQ2; Нория НС-А.20.09 (поз. 3); лист 4 *)
    DI_N3_DP            : BOOL; (* A1 I17 [X17] Датчик подпора; 2SQ3; Нория НС-А.20.09 (поз. 3); лист 4 *)
    DI_N3_SA            : BOOL; (* A1 I18 [X18] Автом./ручн. режим; 2SA1 (11-14); Нория НС-А.20.09 (поз. 3); лист 4 *)
    DI_N3_SB_START      : BOOL; (* A1 I19 [X19] Местный "Пуск" вверху; 2SB1 (13-14, НО); Нория НС-А.20.09 (поз. 3); лист 4 *)
    DI_N3_SB_STOP       : BOOL; (* A1 I20 [X20] Местный "Стоп" вверху; 2SB2 (21-22, НЗ); Нория НС-А.20.09 (поз. 3); лист 4 *)
    DI_N3_SB_ESTOP      : BOOL; (* A1 I21 [X21] Аварийный "Стоп" внизу; 2SB3 (1-2, НЗ); Нория НС-А.20.09 (поз. 3); лист 4 *)
    DI_N3_QF            : BOOL; (* A1 I22 [X22] Защита двигателя нории; 2QF1 (доп. контакт 13-14); Нория НС-А.20.09 (поз. 3); лист 4 *)
    DI_B4_DVU           : BOOL; (* A1 I23 [X23] ДВУ бункера (датчик верхнего уровня); 3SL1 / 3K1; ДВУ/ДНУ бункера БО-2 (поз. 4); лист 5 *)
    (* ---- A1.1 TM3DI32K ---- *)
    DI_B4_DNU           : BOOL; (* A1.1 I0 [1X0] ДНУ бункера (опция); 3K2; ДВУ/ДНУ бункера БО-2 (поз. 4); лист 5 *)
    DI_MUZ5_QF          : BOOL; (* A1.1 I1 [1X1] Защита двигателя МУЗ-8М; 4QF1; Машина универсальная зерноочистительная МУЗ-8М (поз. 5); лист 6 *)
    DI_MUZ5FD_SF        : BOOL; (* A1.1 I2 [1X2] Защита ПЧ; 5SF1; Битер МУЗ-8М (поз. 5), ПЧ 5UZ1; лист 7 *)
    DI_MUZ5FD_FAULT     : BOOL; (* A1.1 I3 [1X3] Авария ПЧ; 5UZ1 (реле 1TA/1TB/1TC); Битер МУЗ-8М (поз. 5), ПЧ 5UZ1; лист 7 *)
    DI_MUZ5FD_READY     : BOOL; (* A1.1 I4 [1X4] Готовность/работа ПЧ; 5UZ1 (реле 2TA/2TB/2TC); Битер МУЗ-8М (поз. 5), ПЧ 5UZ1; лист 7 *)
    DI_MUZ5FD_ESTOP     : BOOL; (* A1.1 I5 [1X5] Аварийный "Стоп"; 5SB1; Битер МУЗ-8М (поз. 5), ПЧ 5UZ1; лист 7 *)
    DI_FAN6_QF          : BOOL; (* A1.1 I6 [1X6] Защита двигателя вентилятора; 6QF1; Вентилятор системы аспирации (поз. 6); лист 8 *)
    DI_SL6_DKS          : BOOL; (* A1.1 I7 [1X7] ДКС шлюзового затвора (датчик контроля скорости); 7SR1; Шлюзовый затвор ЗШ-17 системы аспирации (поз. 6); лист 9 *)
    DI_SL6_QF           : BOOL; (* A1.1 I8 [1X8] Защита двигателя шлюзового затвора; 7QF1; Шлюзовый затвор ЗШ-17 системы аспирации (поз. 6); лист 9 *)
    DI_N7_DKS           : BOOL; (* A1.1 I9 [1X9] ДКС; 8SR1; Нория НС-А.20.09 (поз. 7); лист 10 *)
    DI_N7_DSL1          : BOOL; (* A1.1 I10 [1X10] Датчик сбега ленты 1; 8SQ1; Нория НС-А.20.09 (поз. 7); лист 10 *)
    DI_N7_DSL2          : BOOL; (* A1.1 I11 [1X11] Датчик сбега ленты 2; 8SQ2; Нория НС-А.20.09 (поз. 7); лист 10 *)
    DI_N7_DP            : BOOL; (* A1.1 I12 [1X12] Датчик подпора; 8SQ3; Нория НС-А.20.09 (поз. 7); лист 10 *)
    DI_N7_SA            : BOOL; (* A1.1 I13 [1X13] Автом./ручн. режим; 8SA1; Нория НС-А.20.09 (поз. 7); лист 10 *)
    DI_N7_SB_START      : BOOL; (* A1.1 I14 [1X14] Местный "Пуск" (в заголовке: "вверху"); 8SB1; Нория НС-А.20.09 (поз. 7); лист 10 *)
    DI_N7_SB_STOP       : BOOL; (* A1.1 I15 [1X15] Местный/аварийный "Стоп" на посту внизу (в заголовке: «Местный Стоп вверху»); 8SB2; Нория НС-А.20.09 (поз. 7); лист 10 *)
    DI_N7_SB_ESTOP      : BOOL; (* A1.1 I16 [1X16] Местный стоп нории (вверху) (в заголовке: «Аварийный Стоп внизу»); 8SB3; Нория НС-А.20.09 (поз. 7); лист 10 *)
    DI_N7_QF            : BOOL; (* A1.1 I17 [1X17] Защита двигателя нории; 8QF1; Нория НС-А.20.09 (поз. 7); лист 10 *)
    DI_B8_DVU           : BOOL; (* A1.1 I18 [1X18] ДВУ бункера; 9SL1 / 9K1; ДВУ/ДНУ бункера БО-1 (поз. 8); лист 11 *)
    DI_B8_DNU           : BOOL; (* A1.1 I19 [1X19] ДНУ бункера (опция); 9K2; ДВУ/ДНУ бункера БО-1 (поз. 8); лист 11 *)
    DI_TOR9_QF          : BOOL; (* A1.1 I20 [1X20] Защита двигателя ТОР-18 (на чертеже подписано «Защита двигателя МУЗ-8М» — ошибка копирования); 10QF1; Машина тонкой очистки ТОР-18 (поз. 9); лист 12 *)
    DI_TOR9FD_SF        : BOOL; (* A1.1 I21 [1X21] Защита ПЧ; 11SF1; Машина тонкой очистки ТОР-18 (поз. 9), ПЧ 11UZ1; лист 13 *)
    DI_TOR9FD_FAULT     : BOOL; (* A1.1 I22 [1X22] Авария ПЧ; 11UZ1 (реле 1TA/1TB/1TC); Машина тонкой очистки ТОР-18 (поз. 9), ПЧ 11UZ1; лист 13 *)
    DI_TOR9FD_READY     : BOOL; (* A1.1 I23 [1X23] Готовность/работа ПЧ; 11UZ1 (реле 2TA/2TB/2TC); Машина тонкой очистки ТОР-18 (поз. 9), ПЧ 11UZ1; лист 13 *)
    DI_TOR9FD_ESTOP     : BOOL; (* A1.1 I24 [1X24] Аварийный "Стоп"; 11SB1; Машина тонкой очистки ТОР-18 (поз. 9), ПЧ 11UZ1; лист 13 *)
    DI_FAN10_QF         : BOOL; (* A1.1 I25 [1X25] Защита двигателя вентилятора; 12QF1; Вентилятор системы аспирации (поз. 10); лист 14 *)
    DI_SL10_DKS         : BOOL; (* A1.1 I26 [1X26] ДКС шлюзового затвора; 13SR1; Шлюзовый затвор ЗШ-17 системы аспирации (поз. 10); лист 15 *)
    DI_SL10_QF          : BOOL; (* A1.1 I27 [1X27] Защита двигателя шлюзового затвора; 13QF1; Шлюзовый затвор ЗШ-17 системы аспирации (поз. 10); лист 15 *)
    DI_N11_DKS          : BOOL; (* A1.1 I28 [1X28] ДКС; 14SR1; Нория НС-А.20.09 (поз. 11); лист 16 *)
    DI_N11_DSL1         : BOOL; (* A1.1 I29 [1X29] Датчик сбега ленты 1; 14SQ1; Нория НС-А.20.09 (поз. 11); лист 16 *)
    DI_N11_DSL2         : BOOL; (* A1.1 I30 [1X30] Датчик сбега ленты 2; 14SQ2; Нория НС-А.20.09 (поз. 11); лист 16 *)
    DI_N11_DP           : BOOL; (* A1.1 I31 [1X31] Датчик подпора; 14SQ3; Нория НС-А.20.09 (поз. 11); лист 16 *)
    (* ---- A1.2 TM3DI32K ---- *)
    DI_N11_SA           : BOOL; (* A1.2 I0 [2X0] Автом./ручн. режим; 14SA1; Нория НС-А.20.09 (поз. 11); лист 16 *)
    DI_N11_SB_START     : BOOL; (* A1.2 I1 [2X1] Местный "Пуск" (в заголовке: «вверху»); 14SB1; Нория НС-А.20.09 (поз. 11); лист 16 *)
    DI_N11_SB_STOP      : BOOL; (* A1.2 I2 [2X2] Стоп-грибок на посту внизу (в заголовке: «Местный Стоп вверху»); 14SB2; Нория НС-А.20.09 (поз. 11); лист 16 *)
    DI_N11_SB_ESTOP     : BOOL; (* A1.2 I3 [2X3] Местный стоп нории (вверху) (в заголовке: «Аварийный Стоп внизу»); 14SB3; Нория НС-А.20.09 (поз. 11); лист 16 *)
    DI_N11_QF           : BOOL; (* A1.2 I4 [2X4] Защита двигателя нории; 14QF1; Нория НС-А.20.09 (поз. 11); лист 16 *)
    DI_V121_SF          : BOOL; (* A1.2 I5 [2X5] Защита двигателя переключателя потока; 15SF1; Переключатель потока ППМ-2.160-0/45 (поз. 12.1); лист 17 *)
    DI_V121_POS1        : BOOL; (* A1.2 I6 [2X6] Датчик положения 1 (поток на поз. 13.1); 15SQ1; Переключатель потока ППМ-2.160-0/45 (поз. 12.1); лист 17 *)
    DI_V121_POS2        : BOOL; (* A1.2 I7 [2X7] Датчик положения 2 (поток на поз. 12.2); 15SQ2; Переключатель потока ППМ-2.160-0/45 (поз. 12.1); лист 17 *)
    DI_V122_SF          : BOOL; (* A1.2 I8 [2X8] Защита двигателя переключателя потока; 16SF1; Переключатель потока ППМ-2.160-0/45 (поз. 12.2); лист 18 *)
    DI_V122_POS1        : BOOL; (* A1.2 I9 [2X9] Датчик положения 1 (поток на поз. 14); 16SQ1; Переключатель потока ППМ-2.160-0/45 (поз. 12.2); лист 18 *)
    DI_V122_POS2        : BOOL; (* A1.2 I10 [2X10] Датчик положения 2 (поток на поз. 15.1); 16SQ2; Переключатель потока ППМ-2.160-0/45 (поз. 12.2); лист 18 *)
    DI_V123_SF          : BOOL; (* A1.2 I11 [2X11] Защита двигателя переключателя потока; 17SF1; Переключатель потока ППМ-2.160-0/45 (поз. 12.3); лист 19 *)
    DI_V123_POS1        : BOOL; (* A1.2 I12 [2X12] Датчик положения 1 (поток на поз. 17); 17SQ1; Переключатель потока ППМ-2.160-0/45 (поз. 12.3); лист 19 *)
    DI_V123_POS2        : BOOL; (* A1.2 I13 [2X13] Датчик положения 2 (поток на поз. 20); 17SQ2; Переключатель потока ППМ-2.160-0/45 (поз. 12.3); лист 19 *)
    DI_V124_SF          : BOOL; (* A1.2 I14 [2X14] Защита двигателя переключателя потока; 18SF1; Переключатель потока ППМ-2.160-0/45 (поз. 12.4); лист 20 *)
    DI_V124_POS1        : BOOL; (* A1.2 I15 [2X15] Датчик положения 1 (поток на поз. 22); 18SQ1; Переключатель потока ППМ-2.160-0/45 (поз. 12.4); лист 20 *)
    DI_V124_POS2        : BOOL; (* A1.2 I16 [2X16] Датчик положения 2 (поток на поз. 26); 18SQ2; Переключатель потока ППМ-2.160-0/45 (поз. 12.4); лист 20 *)
    DI_T131_SF          : BOOL; (* A1.2 I17 [2X17] Защита питания ПУ станции затаривания TORBA-1000-1.0 (поз. 13.1); 20SF1; Станция затаривания TORBA-1000-1.0 (поз. 13.1); лист 22 *)
    DI_T132_SF          : BOOL; (* A1.2 I18 [2X18] Защита питания ПУ станции затаривания TORBA-1000-1.0 (поз. 13.2); 21SF1; Станция затаривания TORBA-1000-1.0 (поз. 13.2); лист 22 *)
    DI_T131_DVU         : BOOL; (* A1.2 I19 [2X19] ДВУ бункера TORBA-1000-1.0 (поз. 13.1); 22SL1 / 22K1; Бункер станции затаривания TORBA-1000-1.0 (поз. 13.1); лист 23 *)
    DI_T131_DNU         : BOOL; (* A1.2 I20 [2X20] ДНУ бункера TORBA-1000-1.0 (поз. 13.1); 22SL2 / 22K2; Бункер станции затаривания TORBA-1000-1.0 (поз. 13.1); лист 23 *)
    DI_T132_DVU         : BOOL; (* A1.2 I21 [2X21] ДВУ бункера TORBA-1000-1.0 (поз. 13.2); 23SL1 / 23K1; Бункер станции затаривания TORBA-1000-1.0 (поз. 13.2); лист 24 *)
    DI_T132_DNU         : BOOL; (* A1.2 I22 [2X22] ДНУ бункера TORBA-1000-1.0 (поз. 13.2); 23SL2 / 23K2; Бункер станции затаривания TORBA-1000-1.0 (поз. 13.2); лист 24 *)
    DI_BT141_SF         : BOOL; (* A1.2 I23 [2X23] Защита 1 ПЧ триерного блока; 24SF1; Двигатель 1 триерного блока БТ-9/2 (поз. 14); лист 25 *)
    DI_BT141_FAULT      : BOOL; (* A1.2 I24 [2X24] Авария ПЧ; 24UZ1 (реле 1TA/1TB); Двигатель 1 триерного блока БТ-9/2 (поз. 14); лист 25 *)
    DI_BT141_READY      : BOOL; (* A1.2 I25 [2X25] Готовность/работа ПЧ; 24UZ1 (реле 2TA/2TB); Двигатель 1 триерного блока БТ-9/2 (поз. 14); лист 25 *)
    DI_BT14_ESTOP       : BOOL; (* A1.2 I26 [2X26] Аварийный "Стоп"; 24SB1; Двигатель 1 триерного блока БТ-9/2 (поз. 14); лист 25 *)
    DI_BT142_SF         : BOOL; (* A1.2 I27 [2X27] Защита 2 ПЧ триерного блока; 25SF1; Двигатель 2 триерного блока БТ-9/2 (поз. 14); лист 26 *)
    DI_BT142_FAULT      : BOOL; (* A1.2 I28 [2X28] Авария ПЧ; 25UZ1 (реле 1TA/1TB); Двигатель 2 триерного блока БТ-9/2 (поз. 14); лист 26 *)
    DI_BT142_READY      : BOOL; (* A1.2 I29 [2X29] Готовность/работа ПЧ; 25UZ1 (реле 2TA/2TB); Двигатель 2 триерного блока БТ-9/2 (поз. 14); лист 26 *)
    DI_N16_DKS          : BOOL; (* A1.2 I30 [2X30] ДКС (датчик контроля скорости); 26SR1; Нория НС-А.20.09 (поз. 16); лист 27 *)
    DI_N16_DSL1         : BOOL; (* A1.2 I31 [2X31] Датчик сбега ленты 1; 26SQ1; Нория НС-А.20.09 (поз. 16); лист 27 *)
    (* ---- A1.3 TM3DI32K ---- *)
    DI_N16_DSL2         : BOOL; (* A1.3 I0 [3X0] Датчик сбега ленты 2; 26SQ2; Нория НС-А.20.09 (поз. 16); лист 27 *)
    DI_N16_DP           : BOOL; (* A1.3 I1 [3X1] Датчик подпора; 26SQ3; Нория НС-А.20.09 (поз. 16); лист 27 *)
    DI_N16_SA           : BOOL; (* A1.3 I2 [3X2] Автом./ручн. режим; 26SA1; Нория НС-А.20.09 (поз. 16); лист 27 *)
    DI_N16_SB_START     : BOOL; (* A1.3 I3 [3X3] Местный "Пуск" вверху; 26SB1; Нория НС-А.20.09 (поз. 16); лист 27 *)
    DI_N16_SB_STOP      : BOOL; (* A1.3 I4 [3X4] Местный "Стоп" вверху; 26SB2; Нория НС-А.20.09 (поз. 16); лист 27 *)
    DI_N16_SB_ESTOP     : BOOL; (* A1.3 I5 [3X5] Аварийный "Стоп" внизу; 26SB3; Нория НС-А.20.09 (поз. 16); лист 27 *)
    DI_N16_QF           : BOOL; (* A1.3 I6 [3X6] Защита двигателя нории; 26QF1; Нория НС-А.20.09 (поз. 16); лист 27 *)
    DI_B17_DVU          : BOOL; (* A1.3 I7 [3X7] ДВУ бункера (датчик верхнего уровня); 27SL1 (через реле 27K1); Бункер БО-2 (поз. 17); лист 28 *)
    DI_B17_DNU          : BOOL; (* A1.3 I8 [3X8] ДНУ бункера (опция) (датчик нижнего уровня); 27K2; Бункер БО-2 (поз. 17); лист 28 *)
    DI_KSP18_QF         : BOOL; (* A1.3 I9 [3X9] Защита двигателя КСП-11М; 28QF1; Машина универсальная зерноочистительная КСП-11М (поз. 18); лист 29 *)
    DI_KSP18FD_SF       : BOOL; (* A1.3 I10 [3X10] Защита ПЧ; 29SF1; Машина универсальная зерноочистительная КСП-11М (поз. 18), битер; лист 30 *)
    DI_KSP18FD_FAULT    : BOOL; (* A1.3 I11 [3X11] Авария ПЧ; 29UZ1 (реле 1TA/1TB); Машина универсальная зерноочистительная КСП-11М (поз. 18), битер; лист 30 *)
    DI_KSP18FD_READY    : BOOL; (* A1.3 I12 [3X12] Готовность/работа ПЧ; 29UZ1 (реле 2TA/2TB); Машина универсальная зерноочистительная КСП-11М (поз. 18), битер; лист 30 *)
    DI_KSP18FD_ESTOP    : BOOL; (* A1.3 I13 [3X13] Аварийный "Стоп"; 29SB1; Машина универсальная зерноочистительная КСП-11М (поз. 18); лист 30 *)
    DI_FAN19_QF         : BOOL; (* A1.3 I14 [3X14] Защита двигателя вентилятора; 30QF1; Вентилятор системы аспирации (поз. 19); лист 31 *)
    DI_SL19_DKS         : BOOL; (* A1.3 I15 [3X15] ДКС шлюзового затвора; 31SR1; Шлюзовый затвор ЗШ-17 системы аспирации (поз. 19); лист 32 *)
    DI_SL19_QF          : BOOL; (* A1.3 I16 [3X16] Защита двигателя шлюзового затвора; 31QF1; Шлюзовый затвор ЗШ-17 системы аспирации (поз. 19); лист 32 *)
    DI_N20_DKS          : BOOL; (* A1.3 I17 [3X17] ДКС (датчик контроля скорости); 32SR1; Нория НС-А.20.08 (поз. 20); лист 33 *)
    DI_N20_DSL1         : BOOL; (* A1.3 I18 [3X18] Датчик сбега ленты 1; 32SQ1; Нория НС-А.20.08 (поз. 20); лист 33 *)
    DI_N20_DSL2         : BOOL; (* A1.3 I19 [3X19] Датчик сбега ленты 2; 32SQ2; Нория НС-А.20.08 (поз. 20); лист 33 *)
    DI_N20_DP           : BOOL; (* A1.3 I20 [3X20] Датчик подпора; 32SQ3; Нория НС-А.20.08 (поз. 20); лист 33 *)
    DI_N20_SA           : BOOL; (* A1.3 I21 [3X21] Автом./ручн. режим; 32SA1; Нория НС-А.20.08 (поз. 20); лист 33 *)
    DI_N20_SB_START     : BOOL; (* A1.3 I22 [3X22] Местный "Пуск" вверху; 32SB1; Нория НС-А.20.08 (поз. 20); лист 33 *)
    DI_N20_SB_STOP      : BOOL; (* A1.3 I23 [3X23] Местный "Стоп" вверху; 32SB2; Нория НС-А.20.08 (поз. 20); лист 33 *)
    DI_N20_SB_ESTOP     : BOOL; (* A1.3 I24 [3X24] Аварийный "Стоп" внизу; 32SB3; Нория НС-А.20.08 (поз. 20); лист 33 *)
    DI_N20_QF           : BOOL; (* A1.3 I25 [3X25] Защита двигателя нории; 32QF1; Нория НС-А.20.08 (поз. 20); лист 33 *)
    DI_N21_DKS          : BOOL; (* A1.3 I26 [3X26] ДКС (датчик контроля скорости); 33SR1; Нория НС-А.20.08 (поз. 21); лист 34 *)
    DI_N21_DSL1         : BOOL; (* A1.3 I27 [3X27] Датчик сбега ленты 1; 33SQ1; Нория НС-А.20.08 (поз. 21); лист 34 *)
    DI_N21_DSL2         : BOOL; (* A1.3 I28 [3X28] Датчик сбега ленты 2; 33SQ2; Нория НС-А.20.08 (поз. 21); лист 34 *)
    DI_N21_DP           : BOOL; (* A1.3 I29 [3X29] Датчик подпора; 33SQ3; Нория НС-А.20.08 (поз. 21); лист 34 *)
    DI_N21_SA           : BOOL; (* A1.3 I30 [3X30] Автом./ручн. режим; 33SA1; Нория НС-А.20.08 (поз. 21); лист 34 *)
    DI_N21_SB_START     : BOOL; (* A1.3 I31 [3X31] Местный "Пуск" вверху; 33SB1; Нория НС-А.20.08 (поз. 21); лист 34 *)
    (* ---- A1.4 TM3DI32K ---- *)
    DI_N21_SB_STOP      : BOOL; (* A1.4 I0 [4X0] Местный "Стоп" вверху; 33SB2; Нория НС-А.20.08 (поз. 21); лист 34 *)
    DI_N21_SB_ESTOP     : BOOL; (* A1.4 I1 [4X1] Аварийный "Стоп" внизу; 33SB3; Нория НС-А.20.08 (поз. 21); лист 34 *)
    DI_N21_QF           : BOOL; (* A1.4 I2 [4X2] Защита двигателя нории; 33QF1; Нория НС-А.20.08 (поз. 21); лист 34 *)
    DI_B22_DVU          : BOOL; (* A1.4 I3 [4X3] ДВУ бункера (датчик верхнего уровня); 34SL1 (через реле 34K1); Бункер БО-1 (поз. 22); лист 35 *)
    DI_B22_DNU          : BOOL; (* A1.4 I4 [4X4] ДНУ бункера (опция) (датчик нижнего уровня); 34K2; Бункер БО-1 (поз. 22); лист 35 *)
    DI_SP24FAN_QF       : BOOL; (* A1.4 I5 [4X5] Защита двигателя вентилятора; 35QF1; Стол пневмосортировальный СП-200 (поз. 24), вентилятор; лист 36 *)
    DI_SP24DRV_SF       : BOOL; (* A1.4 I6 [4X6] Защита ПЧ; 36SF1; Стол пневмосортировальный СП-200 (поз. 24), привод стола (ПЧ); лист 37 *)
    DI_SP24DRV_FAULT    : BOOL; (* A1.4 I7 [4X7] Авария ПЧ; 36UZ1 (реле 1TA/1TB); Стол пневмосортировальный СП-200 (поз. 24), привод стола (ПЧ); лист 37 *)
    DI_SP24DRV_READY    : BOOL; (* A1.4 I8 [4X8] Готовность/работа ПЧ; 36UZ1 (реле 2TA/2TB); Стол пневмосортировальный СП-200 (поз. 24), привод стола (ПЧ); лист 37 *)
    DI_SP24DRV_ESTOP    : BOOL; (* A1.4 I9 [4X9] Аварийный "Стоп"; 36SB1; Стол пневмосортировальный СП-200 (поз. 24); лист 37 *)
    DI_FAN25_QF         : BOOL; (* A1.4 I10 [4X10] Защита двигателя вентилятора; 37QF1; Вентилятор системы аспирации (поз. 25); лист 38 *)
    DI_SL25_DKS         : BOOL; (* A1.4 I11 [4X11] ДКС шлюзового затвора; 38SR1; Шлюзовый затвор ЗШ-17 системы аспирации (поз. 25); лист 39 *)
    DI_SL25_QF          : BOOL; (* A1.4 I12 [4X12] Защита двигателя шлюзового затвора; 38QF1; Шлюзовый затвор ЗШ-17 системы аспирации (поз. 25); лист 39 *)
    DI_FAN28_QF         : BOOL; (* A1.4 I13 [4X13] Защита двигателя вентилятора; 39QF1; Вентилятор системы аспирации (поз. 28); лист 40 *)
    DI_SL28_DKS         : BOOL; (* A1.4 I14 [4X14] ДКС шлюзового затвора; 40SR1; Шлюзовый затвор ЗШ-17 системы аспирации (поз. 28); лист 41 *)
    DI_SL28_QF          : BOOL; (* A1.4 I15 [4X15] Защита двигателя шлюзового затвора; 40QF1; Шлюзовый затвор ЗШ-17 системы аспирации (поз. 28); лист 41 *)
    DI_SH31_DKS         : BOOL; (* A1.4 I16 [4X16] ДКС (датчик контроля скорости); 41SR1; Конвейер шнековый КШУ-150 5,5М/5 (поз. 31); лист 42 *)
    DI_SH31_DP          : BOOL; (* A1.4 I17 [4X17] Датчик подпора; 41SQ1; Конвейер шнековый КШУ-150 5,5М/5 (поз. 31); лист 42 *)
    DI_SH31_SA          : BOOL; (* A1.4 I18 [4X18] Автом./ручн. режим; 41SA1; Конвейер шнековый КШУ-150 5,5М/5 (поз. 31); лист 42 *)
    DI_SH31_SB_START    : BOOL; (* A1.4 I19 [4X19] Местный "Пуск"; 41SB1; Конвейер шнековый КШУ-150 5,5М/5 (поз. 31); лист 42 *)
    DI_SH31_SB_STOP     : BOOL; (* A1.4 I20 [4X20] Местный "Стоп"; 41SB2; Конвейер шнековый КШУ-150 5,5М/5 (поз. 31); лист 42 *)
    DI_SH31_SB_END      : BOOL; (* A1.4 I21 [4X21] Местный "Стоп" в конце конвейера; 41SB3; Конвейер шнековый КШУ-150 5,5М/5 (поз. 31); лист 42 *)
    DI_SH31_QF          : BOOL; (* A1.4 I22 [4X22] Защита двигателя конвейера; 41QF1; Конвейер шнековый КШУ-150 5,5М/5 (поз. 31); лист 42 *)
    DI_SH32_DKS         : BOOL; (* A1.4 I23 [4X23] ДКС (датчик контроля скорости); 42SR1; Конвейер шнековый КШУ-150 6М/5 (поз. 32); лист 43 *)
    DI_SH32_DP          : BOOL; (* A1.4 I24 [4X24] Датчик подпора; 42SQ1; Конвейер шнековый КШУ-150 6М/5 (поз. 32); лист 43 *)
    DI_SH32_SA          : BOOL; (* A1.4 I25 [4X25] Автом./ручн. режим; 42SA1; Конвейер шнековый КШУ-150 6М/5 (поз. 32); лист 43 *)
    DI_SH32_SB_START    : BOOL; (* A1.4 I26 [4X26] Местный "Пуск"; 42SB1; Конвейер шнековый КШУ-150 6М/5 (поз. 32); лист 43 *)
    DI_SH32_SB_STOP     : BOOL; (* A1.4 I27 [4X27] Местный "Стоп"; 42SB2; Конвейер шнековый КШУ-150 6М/5 (поз. 32); лист 43 *)
    DI_SH32_SB_END      : BOOL; (* A1.4 I28 [4X28] Местный "Стоп" в конце конвейера; 42SB3; Конвейер шнековый КШУ-150 6М/5 (поз. 32); лист 43 *)
    DI_SH32_QF          : BOOL; (* A1.4 I29 [4X29] Защита двигателя конвейера; 42QF1; Конвейер шнековый КШУ-150 6М/5 (поз. 32); лист 43 *)
    DI_SH33_DKS         : BOOL; (* A1.4 I30 [4X30] ДКС (датчик контроля скорости); 43SR1; Конвейер шнековый КШУ-150 6М/5 (поз. 33); лист 44 *)
    DI_SH33_DP          : BOOL; (* A1.4 I31 [4X31] Датчик подпора; 43SQ1; Конвейер шнековый КШУ-150 6М/5 (поз. 33); лист 44 *)
    (* ---- A1.5 TM3DI32K ---- *)
    DI_SH33_SA          : BOOL; (* A1.5 I0 [5X0] Автом./ручн. режим; 43SA1; Конвейер шнековый КШУ-150 6М/5 (поз. 33); лист 44 *)
    DI_SH33_SB_START    : BOOL; (* A1.5 I1 [5X1] Местный "Пуск"; 43SB1; Конвейер шнековый КШУ-150 6М/5 (поз. 33); лист 44 *)
    DI_SH33_SB_STOP     : BOOL; (* A1.5 I2 [5X2] Местный "Стоп"; 43SB2; Конвейер шнековый КШУ-150 6М/5 (поз. 33); лист 44 *)
    DI_SH33_SB_END      : BOOL; (* A1.5 I3 [5X3] Местный "Стоп" в конце конвейера; 43SB3; Конвейер шнековый КШУ-150 6М/5 (поз. 33); лист 44 *)
    DI_SH33_QF          : BOOL; (* A1.5 I4 [5X4] Защита двигателя конвейера; 43QF1; Конвейер шнековый КШУ-150 6М/5 (поз. 33); лист 44 *)
    DI_KC34_DKS         : BOOL; (* A1.5 I5 [5X5] ДКС (датчик контроля скорости); 44KM2 (от РДД-03); Конвейер цепной КЦСВ (поз. 34); лист 45 *)
    DI_KC34_DP          : BOOL; (* A1.5 I6 [5X6] Датчик подпора; 44KM3 (от РСУ-4); Конвейер цепной КЦСВ (поз. 34); лист 45 *)
    DI_KC34_SA          : BOOL; (* A1.5 I7 [5X7] Автом./ручн. режим; 44SA1; Конвейер цепной КЦСВ (поз. 34); лист 45 *)
    DI_KC34_SB_START    : BOOL; (* A1.5 I8 [5X8] Местный "Пуск"; 44SB1; Конвейер цепной КЦСВ (поз. 34); лист 45 *)
    DI_KC34_SB_STOP     : BOOL; (* A1.5 I9 [5X9] Местный "Стоп"; 44SB2; Конвейер цепной КЦСВ (поз. 34); лист 45 *)
    DI_KC34_SB_END      : BOOL; (* A1.5 I10 [5X10] Местный "Стоп" в конце конвейера; 44SB3; Конвейер цепной КЦСВ (поз. 34); лист 45 *)
    DI_KC34_QF          : BOOL; (* A1.5 I11 [5X11] Защита двигателя конвейера; 44QF1; Конвейер цепной КЦСВ (поз. 34); лист 45 *)
    DI_KC35_DKS         : BOOL; (* A1.5 I12 [5X12] ДКС; 45KM2 (контакт 13-14); Конвейер цепной КЦСН (поз. 35); лист 47 *)
    DI_KC35_DP          : BOOL; (* A1.5 I13 [5X13] Датчик подпора; 45KM3 (контакт 13-14); Конвейер цепной КЦСН (поз. 35); лист 47 *)
    DI_KC35_SA          : BOOL; (* A1.5 I14 [5X14] Автом./ручн. режим; 45SA1 (13-14); Конвейер цепной КЦСН (поз. 35); лист 47 *)
    DI_KC35_SB_START    : BOOL; (* A1.5 I15 [5X15] Местный "Пуск"; 45SB1 (13-14, НО); Конвейер цепной КЦСН (поз. 35); лист 47 *)
    DI_KC35_SB_STOP     : BOOL; (* A1.5 I16 [5X16] Местный "Стоп"; 45SB2 (21-22, НЗ); Конвейер цепной КЦСН (поз. 35); лист 47 *)
    DI_KC35_SB_END      : BOOL; (* A1.5 I17 [5X17] Местный "Стоп" в конце конвейера; 45SB3, 45SB4 (1-2, НЗ, последовательно); Конвейер цепной КЦСН (поз. 35); лист 47 *)
    DI_KC35_QF          : BOOL; (* A1.5 I18 [5X18] Защита двигателя конвейера; 45QF1 (доп. контакт 13-14); Конвейер цепной КЦСН (поз. 35); лист 47 *)
    DI_KC36_DKS         : BOOL; (* A1.5 I19 [5X19] ДКС; 46KM2 (контакт 13-14); Конвейер цепной КЦСН (поз. 36); лист 49 *)
    DI_KC36_DP          : BOOL; (* A1.5 I20 [5X20] Датчик подпора; 46KM3 (контакт 13-14); Конвейер цепной КЦСН (поз. 36); лист 49 *)
    DI_KC36_SA          : BOOL; (* A1.5 I21 [5X21] Автом./ручн. режим; 46SA1 (13-14); Конвейер цепной КЦСН (поз. 36); лист 49 *)
    DI_KC36_SB_START    : BOOL; (* A1.5 I22 [5X22] Местный "Пуск"; 46SB1 (13-14, НО); Конвейер цепной КЦСН (поз. 36); лист 49 *)
    DI_KC36_SB_STOP     : BOOL; (* A1.5 I23 [5X23] Местный "Стоп"; 46SB2 (21-22, НЗ); Конвейер цепной КЦСН (поз. 36); лист 49 *)
    DI_KC36_SB_END      : BOOL; (* A1.5 I24 [5X24] Местный "Стоп" в конце конвейера; 46SB3 (1-2, НЗ); Конвейер цепной КЦСН (поз. 36); лист 49 *)
    DI_KC36_QF          : BOOL; (* A1.5 I25 [5X25] Защита двигателя конвейера; 46QF1 (доп. контакт 13-14); Конвейер цепной КЦСН (поз. 36); лист 49 *)
    DI_SH30_DKS         : BOOL; (* A1.5 I26 [5X26] ДКС (опция); — (датчик не указан, клеммная коробка 1-47КО); Конвейер (поз. 30); лист 51 *)
    DI_SH30_DP          : BOOL; (* A1.5 I27 [5X27] Датчик подпора (опция); — (датчик не указан, 1-47КО); Конвейер (поз. 30); лист 51 *)
    DI_SH30_SA          : BOOL; (* A1.5 I28 [5X28] Автом./ручн. режим; 47SA1 (13-14); Конвейер (поз. 30); лист 51 *)
    DI_SH30_SB_START    : BOOL; (* A1.5 I29 [5X29] Местный "Пуск"; 47SB1 (13-14, НО); Конвейер (поз. 30); лист 51 *)
    DI_SH30_SB_STOP     : BOOL; (* A1.5 I30 [5X30] Местный "Стоп"; 47SB2 (21-22, НЗ); Конвейер (поз. 30); лист 51 *)
    DI_SH30_SB_END      : BOOL; (* A1.5 I31 [5X31] Местный "Стоп" в конце конвейера; 47SB3 (1-2, НЗ); Конвейер (поз. 30); лист 51 *)
    (* ---- A1.6 TM3DI32K ---- *)
    DI_SH30_QF          : BOOL; (* A1.6 I0 [6X0] Защита двигателя конвейера; 47QF1 (доп. контакт 13-14); Конвейер (поз. 30); лист 51 *)
    DI_ZN26_DKS         : BOOL; (* A1.6 I1 [6X1] ДКС; 48SR1; Нория зерновая 5КТ-20 тип Z (поз. 26); лист 53 *)
    DI_ZN26_RES         : BOOL; (* A1.6 I2 [6X2] Резерв; —; Нория зерновая 5КТ-20 тип Z (поз. 26); лист 53 *)
    DI_ZN26_SA          : BOOL; (* A1.6 I3 [6X3] Автом./ручн. режим; 48SA1 (13-14); Нория зерновая 5КТ-20 тип Z (поз. 26); лист 53 *)
    DI_ZN26_SB_START    : BOOL; (* A1.6 I4 [6X4] Местный "Пуск"; 48SB1 (13-14, НО); Нория зерновая 5КТ-20 тип Z (поз. 26); лист 53 *)
    DI_ZN26_SB_STOP     : BOOL; (* A1.6 I5 [6X5] Местный "Стоп"; 48SB2 (21-22, НЗ); Нория зерновая 5КТ-20 тип Z (поз. 26); лист 53 *)
    DI_ZN26_SB_END      : BOOL; (* A1.6 I6 [6X6] Местный "Стоп" в конце нории; 48SB3 (1-2, НЗ); Нория зерновая 5КТ-20 тип Z (поз. 26); лист 53 *)
    DI_ZN26_FAULT       : BOOL; (* A1.6 I7 [6X7] Авария ПЧ; 48UZ1 реле 1T (клеммы 1TB-1TA); Нория зерновая 5КТ-20 тип Z (поз. 26); лист 53 *)
    DI_ZN26_READY       : BOOL; (* A1.6 I8 [6X8] Готовность/работа ПЧ; 48UZ1 реле 2T (клеммы 2TB-2TA); Нория зерновая 5КТ-20 тип Z (поз. 26); лист 53 *)
    DI_ZN26_SF          : BOOL; (* A1.6 I9 [6X9] Защита ПЧ; 48SF1 (доп. контакт 13-14); Нория зерновая 5КТ-20 тип Z (поз. 26); лист 53 *)
    DI_V49_ON           : BOOL; (* A1.6 I10 [6X10] Механизм выгрузки включен; 49SQ1 (11-12); Промежуточная выгрузка нории (поз. 26) — поток на TORBA-1000 (поз. 13.2); лист 54 *)
    DI_V49_OFF          : BOOL; (* A1.6 I11 [6X11] Механизм выгрузки выключен; 49SQ2 (11-12); Промежуточная выгрузка нории (поз. 26) — поток на TORBA-1000 (поз. 13.2); лист 54 *)
    DI_ZN29_DKS         : BOOL; (* A1.6 I12 [6X12] ДКС; 50SR1; Нория зерновая 5КТ-20 тип Z (поз. 29); лист 56 *)
    DI_ZN29_RES         : BOOL; (* A1.6 I13 [6X13] Резерв; —; Нория зерновая 5КТ-20 тип Z (поз. 29); лист 56 *)
    DI_ZN29_SA          : BOOL; (* A1.6 I14 [6X14] Автом./ручн. режим; 50SA1 (13-14); Нория зерновая 5КТ-20 тип Z (поз. 29); лист 56 *)
    DI_ZN29_SB_START    : BOOL; (* A1.6 I15 [6X15] Местный "Пуск"; 50SB1 (13-14, НО); Нория зерновая 5КТ-20 тип Z (поз. 29); лист 56 *)
    DI_ZN29_SB_STOP     : BOOL; (* A1.6 I16 [6X16] Местный "Стоп"; 50SB2 (21-22, НЗ); Нория зерновая 5КТ-20 тип Z (поз. 29); лист 56 *)
    DI_ZN29_SB_END      : BOOL; (* A1.6 I17 [6X17] Местный "Стоп" в конце нории; 50SB3 (1-2, НЗ); Нория зерновая 5КТ-20 тип Z (поз. 29); лист 56 *)
    DI_ZN29_FAULT       : BOOL; (* A1.6 I18 [6X18] Авария ПЧ; 50UZ1 реле 1T (1TB-1TA); Нория зерновая 5КТ-20 тип Z (поз. 29); лист 56 *)
    DI_ZN29_READY       : BOOL; (* A1.6 I19 [6X19] Готовность/работа ПЧ; 50UZ1 реле 2T (2TB-2TA); Нория зерновая 5КТ-20 тип Z (поз. 29); лист 56 *)
    DI_ZN29_SF          : BOOL; (* A1.6 I20 [6X20] Защита ПЧ; 50SF1 (доп. контакт 13-14); Нория зерновая 5КТ-20 тип Z (поз. 29); лист 56 *)
    DI_GATE1_OPENED     : BOOL; (* A1.6 I21 [6X21] Открыта заслонка; 51SQ1; Заслонка (поз. 1); лист 58 *)
    DI_GATE1_CLOSED     : BOOL; (* A1.6 I22 [6X22] Закрыта заслонка; 51SQ2; Заслонка (поз. 1); лист 58 *)
    DI_GATE1_SA         : BOOL; (* A1.6 I23 [6X23] Автом./ручн. режим; 51SA1 (13-14); Заслонка (поз. 1); лист 58 *)
    DI_GATE1_SB_OPEN    : BOOL; (* A1.6 I24 [6X24] Открыть заслонку; 51SB1 (13-14, НО); Заслонка (поз. 1); лист 58 *)
    DI_GATE1_SB_CLOSE   : BOOL; (* A1.6 I25 [6X25] Закрыть заслонку; 51SB2 (13-14, НО); Заслонка (поз. 1); лист 58 *)
    DI_GATE1_SB_STOP    : BOOL; (* A1.6 I26 [6X26] Местный "Стоп"; 51SB3 (1-2, НЗ); Заслонка (поз. 1); лист 58 *)
    DI_GATE1_FAULT      : BOOL; (* A1.6 I27 [6X27] Авария ПЧ; 51UZ1 реле 1T (1TB-1TA); Заслонка (поз. 1); лист 58 *)
    DI_GATE1_READY      : BOOL; (* A1.6 I28 [6X28] Готовность/работа ПЧ; 51UZ1 реле 2T (2TB-2TA); Заслонка (поз. 1); лист 58 *)
    DI_GATE1_SF         : BOOL; (* A1.6 I29 [6X29] Защита ПЧ; 51SF1 (доп. контакт 13-14); Заслонка (поз. 1); лист 58 *)
    DI_B27_DVU1         : BOOL; (* A1.6 I30 [6X30] ДВУ бункера; 52SL1 через реле 52K1 (11-14); ДВУ бункера (поз. 27); лист 59 *)
    DI_B27_DVU2         : BOOL; (* A1.6 I31 [6X31] ДВУ бункера; 52SL2 через реле 52K2 (11-14); ДВУ бункера (поз. 27); лист 59 *)
    (* ---- A1.7 TM3DI32K ---- *)
    DI_FS27_ASP_SF      : BOOL; (* A1.7 I0 [7X0] Защита питания аспирации; 53SF1 (доп. контакт 11-14); Питание аспирации (поз. 27) — опция; лист 60 *)
    DI_FS27_SF          : BOOL; (* A1.7 I1 [7X1] Защита питания фотосепаратора; 54SF1 (доп. контакт 11-14); Питание фотосепаратора (поз. 27); лист 60 *)
    DI_FS27_STATUS      : BOOL; (* A1.7 I2 [7X2] Статус аппарата; Фотосепаратор, выход (O4) =RE-A6-X24:1; Фотоэлектронный сепаратор (поз. 27); лист 61 *)
    DI_FS27_REMOTE      : BOOL; (* A1.7 I3 [7X3] Внешнее управление; Фотосепаратор, выход (O5) =RE-A6-X25:4; Фотоэлектронный сепаратор (поз. 27); лист 61 *)
    DI_FS27_ERROR       : BOOL; (* A1.7 I4 [7X4] Критическая ошибка; Фотосепаратор, выход (O7) =RE-A6-X25:2; Фотоэлектронный сепаратор (поз. 27); лист 61 *)
    DI_DRYER_SF         : BOOL; (* A1.7 I5 [7X5] Защита питания осушителя (опция); 56SF1 (доп. контакт 11-14); Питание осушителя (поз. 45) — опция; лист 62 *)
    DI_COMPR_SF         : BOOL; (* A1.7 I6 [7X6] Защита питания компрессора (поз. 45); 57SF1 (доп. контакт 11-14); Питание компрессора (поз. 45) 15,0кВт 32,0А; лист 62 *)
    DI_COMPR2_SF        : BOOL; (* A1.7 I7 [7X7] Защита питания компрессора (опция); 58SF1 (на схеме у входа), фактически автомат 58QF1 4,0-6,3А; Питание компрессора (опция) 2,2кВт 5,0А; лист 62 *)
    DI_A17_I8_RES       : BOOL; (* A1.7 I8 [7X8] Резерв; 59K3 (11-14); Резерв (интерфейс сухих контактов, клеммы X8); лист 66 *)
    DI_A17_I9_RES       : BOOL; (* A1.7 I9 [7X9] Резерв; 59K4 (11-14); Резерв (интерфейс сухих контактов, клеммы X8); лист 66 *)
    (* ---- A1 TM241CE40T ---- *)
    DO_SIREN            : BOOL; (* A1 Q0 [Y0] Сирена; HAK1; Шкаф управления — общие сигналы; лист 3 *)
    DO_LAMP_ALARM       : BOOL; (* A1 Q1 [Y1] Сигнал "Авария"; HL6; Шкаф управления — общие сигналы; лист 3 *)
    DO_N3_RUN           : BOOL; (* A1 Q2 [Y2] Включение нории; 2K1; Нория НС-А.20.09 (поз. 3); лист 4 *)
    DO_MUZ5_RUN         : BOOL; (* A1 Q3 [Y3] Включить МУЗ-8М; 4K1 / 4KM1; Машина универсальная зерноочистительная МУЗ-8М (поз. 5); лист 6 *)
    DO_MUZ5FD_POWER     : BOOL; (* A1 Q4 [Y4] Включить ПЧ; 5K1 / 5KM1; Битер МУЗ-8М (поз. 5), ПЧ 5UZ1; лист 7 *)
    DO_MUZ5FD_RESET     : BOOL; (* A1 Q5 [Y5] Сброс аварии ПЧ; 5K2; Битер МУЗ-8М (поз. 5), ПЧ 5UZ1; лист 7 *)
    DO_MUZ5FD_RUN       : BOOL; (* A1 Q6 [Y6] Пуск битера; 5K3; Битер МУЗ-8М (поз. 5), ПЧ 5UZ1; лист 7 *)
    DO_FAN6_RUN         : BOOL; (* A1 Q7 [Y7] Включить вентилятор аспирации; 6K1 / 6KM1; Вентилятор системы аспирации (поз. 6); лист 8 *)
    DO_SL6_RUN          : BOOL; (* A1 Q8 [Y8] Включить затвор шлюзовый; 7K1 / 7KM1; Шлюзовый затвор ЗШ-17 системы аспирации (поз. 6); лист 9 *)
    DO_N7_RUN           : BOOL; (* A1 Q9 [Y9] Включение нории; 8K1 / 8KM1; Нория НС-А.20.09 (поз. 7); лист 10 *)
    DO_TOR9_RUN         : BOOL; (* A1 Q10 [Y10] Включить ТОР-18; 10K1 / 10KM1; Машина тонкой очистки ТОР-18 (поз. 9); лист 12 *)
    DO_TOR9FD_POWER     : BOOL; (* A1 Q11 [Y11] Включить ПЧ; 11K1 / 11KM1; Машина тонкой очистки ТОР-18 (поз. 9), ПЧ 11UZ1; лист 13 *)
    DO_TOR9FD_RESET     : BOOL; (* A1 Q12 [Y12] Сброс аварии ПЧ; 11K2; Машина тонкой очистки ТОР-18 (поз. 9), ПЧ 11UZ1; лист 13 *)
    DO_TOR9FD_RUN       : BOOL; (* A1 Q13 [Y13] Пуск (ПЧ ТОР-18); 11K3; Машина тонкой очистки ТОР-18 (поз. 9), ПЧ 11UZ1; лист 13 *)
    DO_FAN10_RUN        : BOOL; (* A1 Q14 [Y14] Включить вентилятор аспирации; 12K1 / 12KM1; Вентилятор системы аспирации (поз. 10); лист 14 *)
    DO_SL10_RUN         : BOOL; (* A1 Q15 [Y15] Включить затвор шлюзовый; 13K1 / 13KM1; Шлюзовый затвор ЗШ-17 системы аспирации (поз. 10); лист 15 *)
    (* ---- A1.8 TM3DQ32TK ---- *)
    DO_N11_RUN          : BOOL; (* A1.8 Q0 [8Y0] Включение нории; 14K1 / 14KM1; Нория НС-А.20.09 (поз. 11); лист 16 *)
    DO_V121_POS1        : BOOL; (* A1.8 Q1 [8Y1] Поток на (поз. 13.1); 15K1; Переключатель потока ППМ-2.160-0/45 (поз. 12.1); лист 17 *)
    DO_V121_POS2        : BOOL; (* A1.8 Q2 [8Y2] Поток на (поз. 12.2); 15K2; Переключатель потока ППМ-2.160-0/45 (поз. 12.1); лист 17 *)
    DO_V122_POS1        : BOOL; (* A1.8 Q3 [8Y3] Поток на (поз. 14); 16K1; Переключатель потока ППМ-2.160-0/45 (поз. 12.2); лист 18 *)
    DO_V122_POS2        : BOOL; (* A1.8 Q4 [8Y4] Поток на (поз. 15.1); 16K2; Переключатель потока ППМ-2.160-0/45 (поз. 12.2); лист 18 *)
    DO_V123_POS1        : BOOL; (* A1.8 Q5 [8Y5] Поток на (поз. 17); 17K1; Переключатель потока ППМ-2.160-0/45 (поз. 12.3); лист 19 *)
    DO_V123_POS2        : BOOL; (* A1.8 Q6 [8Y6] Поток на (поз. 20); 17K2; Переключатель потока ППМ-2.160-0/45 (поз. 12.3); лист 19 *)
    DO_V124_POS1        : BOOL; (* A1.8 Q7 [8Y7] Поток на (поз. 22); 18K1; Переключатель потока ППМ-2.160-0/45 (поз. 12.4); лист 20 *)
    DO_V124_POS2        : BOOL; (* A1.8 Q8 [8Y8] Поток на (поз. 26); 18K2; Переключатель потока ППМ-2.160-0/45 (поз. 12.4); лист 20 *)
    DO_A18_Q9_RES       : BOOL; (* A1.8 Q9 [8Y9] Резерв; 19K1; (лист 21, без заголовка; рядом цепь «Включить питание» 19KM1); лист 21 *)
    DO_BT141_POWER      : BOOL; (* A1.8 Q10 [8Y10] Включить ПЧ; 24K1; Двигатель 1 триерного блока БТ-9/2 (поз. 14); лист 25 *)
    DO_BT141_RESET      : BOOL; (* A1.8 Q11 [8Y11] Сброс аварии ПЧ; 24K2; Двигатель 1 триерного блока БТ-9/2 (поз. 14); лист 25 *)
    DO_BT141_RUN        : BOOL; (* A1.8 Q12 [8Y12] Пуск триера; 24K3; Двигатель 1 триерного блока БТ-9/2 (поз. 14); лист 25 *)
    DO_BT142_POWER      : BOOL; (* A1.8 Q13 [8Y13] Включить ПЧ; 25K1; Двигатель 2 триерного блока БТ-9/2 (поз. 14); лист 26 *)
    DO_BT142_RESET      : BOOL; (* A1.8 Q14 [8Y14] Сброс аварии ПЧ; 25K2; Двигатель 2 триерного блока БТ-9/2 (поз. 14); лист 26 *)
    DO_BT142_RUN        : BOOL; (* A1.8 Q15 [8Y15] Пуск триера; 25K3; Двигатель 2 триерного блока БТ-9/2 (поз. 14); лист 26 *)
    DO_N16_RUN          : BOOL; (* A1.8 Q16 [8Y16] Включение нории; 26K1; Нория НС-А.20.09 (поз. 16); лист 27 *)
    DO_KSP18_RUN        : BOOL; (* A1.8 Q17 [8Y17] Включить КСП-11М; 28K1; Машина универсальная зерноочистительная КСП-11М (поз. 18); лист 29 *)
    DO_KSP18FD_POWER    : BOOL; (* A1.8 Q18 [8Y18] Включить ПЧ; 29K1; Машина универсальная зерноочистительная КСП-11М (поз. 18), битер; лист 30 *)
    DO_KSP18FD_RESET    : BOOL; (* A1.8 Q19 [8Y19] Сброс аварии ПЧ; 29K2; Машина универсальная зерноочистительная КСП-11М (поз. 18), битер; лист 30 *)
    DO_KSP18FD_RUN      : BOOL; (* A1.8 Q20 [8Y20] Пуск битера; 29K3; Машина универсальная зерноочистительная КСП-11М (поз. 18), битер; лист 30 *)
    DO_FAN19_RUN        : BOOL; (* A1.8 Q21 [8Y21] Включить вентилятор аспирации; 30K1; Вентилятор системы аспирации (поз. 19); лист 31 *)
    DO_SL19_RUN         : BOOL; (* A1.8 Q22 [8Y22] Включить затвор шлюзовый; 31K1; Шлюзовый затвор ЗШ-17 системы аспирации (поз. 19); лист 32 *)
    DO_N20_RUN          : BOOL; (* A1.8 Q23 [8Y23] Включение нории; 32K1; Нория НС-А.20.08 (поз. 20); лист 33 *)
    DO_N21_RUN          : BOOL; (* A1.8 Q24 [8Y24] Включение нории; 33K1; Нория НС-А.20.08 (поз. 21); лист 34 *)
    DO_SP24FAN_RUN      : BOOL; (* A1.8 Q25 [8Y25] Включить вентилятор стола СП-200; 35K1; Стол пневмосортировальный СП-200 (поз. 24), вентилятор; лист 36 *)
    DO_SP24DRV_POWER    : BOOL; (* A1.8 Q26 [8Y26] Включить ПЧ; 36K1; Стол пневмосортировальный СП-200 (поз. 24), привод стола (ПЧ); лист 37 *)
    DO_SP24DRV_RESET    : BOOL; (* A1.8 Q27 [8Y27] Сброс аварии ПЧ; 36K2; Стол пневмосортировальный СП-200 (поз. 24), привод стола (ПЧ); лист 37 *)
    DO_SP24DRV_RUN      : BOOL; (* A1.8 Q28 [8Y28] Пуск битера; 36K3; Стол пневмосортировальный СП-200 (поз. 24), привод стола (ПЧ); лист 37 *)
    DO_FAN25_RUN        : BOOL; (* A1.8 Q29 [8Y29] Включить вентилятор аспирации; 37K1; Вентилятор системы аспирации (поз. 25); лист 38 *)
    DO_SL25_RUN         : BOOL; (* A1.8 Q30 [8Y30] Включить затвор шлюзовый; 38K1; Шлюзовый затвор ЗШ-17 системы аспирации (поз. 25); лист 39 *)
    DO_FAN28_RUN        : BOOL; (* A1.8 Q31 [8Y31] Включить вентилятор аспирации; 39K1; Вентилятор системы аспирации (поз. 28); лист 40 *)
    (* ---- A1.9 TM3DQ32TK ---- *)
    DO_SL28_RUN         : BOOL; (* A1.9 Q0 [9Y0] Включить затвор шлюзовый; 40K1; Шлюзовый затвор ЗШ-17 системы аспирации (поз. 28); лист 41 *)
    DO_SH31_RUN         : BOOL; (* A1.9 Q1 [9Y1] Включение конвейера; 41K1; Конвейер шнековый КШУ-150 5,5М/5 (поз. 31); лист 42 *)
    DO_SH32_RUN         : BOOL; (* A1.9 Q2 [9Y2] Включение конвейера; 42K1; Конвейер шнековый КШУ-150 6М/5 (поз. 32); лист 43 *)
    DO_SH33_RUN         : BOOL; (* A1.9 Q3 [9Y3] Включение конвейера; 43K1; Конвейер шнековый КШУ-150 6М/5 (поз. 33); лист 44 *)
    DO_KC34_RUN         : BOOL; (* A1.9 Q4 [9Y4] Включение конвейера; 44K1; Конвейер цепной КЦСВ (поз. 34); лист 45 *)
    DO_KC35_RUN         : BOOL; (* A1.9 Q5 [9Y5] Включение конвейера; 45K1; Конвейер цепной КЦСН (поз. 35); лист 47 *)
    DO_KC36_RUN         : BOOL; (* A1.9 Q6 [9Y6] Включение конвейера; 46K1; Конвейер цепной КЦСН (поз. 36); лист 49 *)
    DO_SH30_RUN         : BOOL; (* A1.9 Q7 [9Y7] Включение конвейера; 47K1; Конвейер (поз. 30); лист 51 *)
    DO_ZN26_POWER       : BOOL; (* A1.9 Q8 [9Y8] Включение ПЧ; 48K1; Нория зерновая 5КТ-20 тип Z (поз. 26); лист 53 *)
    DO_ZN26_RUN         : BOOL; (* A1.9 Q9 [9Y9] Включение нории; 48K2; Нория зерновая 5КТ-20 тип Z (поз. 26); лист 53 *)
    DO_ZN26_RESET       : BOOL; (* A1.9 Q10 [9Y10] Сброс аварии; 48K3; Нория зерновая 5КТ-20 тип Z (поз. 26); лист 53 *)
    DO_V49_ON           : BOOL; (* A1.9 Q11 [9Y11] Включить механизм выгрузки; 49K1; Промежуточная выгрузка нории (поз. 26) — поток на TORBA-1000 (поз. 13.2); лист 54 *)
    DO_V49_OFF          : BOOL; (* A1.9 Q12 [9Y12] Отключить механизм выгрузки; 49K2; Промежуточная выгрузка нории (поз. 26) — поток на TORBA-1000 (поз. 13.2); лист 54 *)
    DO_ZN29_POWER       : BOOL; (* A1.9 Q13 [9Y13] Включение ПЧ; 50K1; Нория зерновая 5КТ-20 тип Z (поз. 29); лист 56 *)
    DO_ZN29_RUN         : BOOL; (* A1.9 Q14 [9Y14] Включение нории; 50K2; Нория зерновая 5КТ-20 тип Z (поз. 29); лист 56 *)
    DO_ZN29_RESET       : BOOL; (* A1.9 Q15 [9Y15] Сброс аварии; 50K3; Нория зерновая 5КТ-20 тип Z (поз. 29); лист 56 *)
    DO_GATE1_POWER      : BOOL; (* A1.9 Q16 [9Y16] Включение ПЧ; 51K1; Заслонка (поз. 1); лист 58 *)
    DO_GATE1_OPEN       : BOOL; (* A1.9 Q17 [9Y17] Открытие заслонки; 51K2; Заслонка (поз. 1); лист 58 *)
    DO_GATE1_RESET      : BOOL; (* A1.9 Q18 [9Y18] Сброс аварии; 51K3; Заслонка (поз. 1); лист 58 *)
    DO_GATE1_CLOSE      : BOOL; (* A1.9 Q19 [9Y19] Закрытие заслонки; 51K5; Заслонка (поз. 1); лист 58 *)
    DO_FS27_ON          : BOOL; (* A1.9 Q20 [9Y20] Включить аппарат; 55K1; Фотоэлектронный сепаратор (поз. 27); лист 61 *)
    DO_FS27_OFF         : BOOL; (* A1.9 Q21 [9Y21] Выключить аппарат; 55K2; Фотоэлектронный сепаратор (поз. 27); лист 61 *)
    DO_FS27_ENABLE      : BOOL; (* A1.9 Q22 [9Y22] Разрешить секцию 1-3; 55K3; Фотоэлектронный сепаратор (поз. 27); лист 61 *)
    DO_A19_Q23_RES      : BOOL; (* A1.9 Q23 [9Y23] Резерв; 59K1; Резерв (интерфейс сухих контактов, клеммы X8); лист 66 *)
    DO_A19_Q24_RES      : BOOL; (* A1.9 Q24 [9Y24] Резерв; 59K2; Резерв (интерфейс сухих контактов, клеммы X8); лист 66 *)
END_VAR

(* global variable list GVL_Retain *)
(* Уставки и моточасы. При необходимости сохранять их и при загрузке новой программы
   перенести эти переменные в список Persistent (VAR_GLOBAL PERSISTENT RETAIN). *)
VAR_GLOBAL RETAIN
    uInitMagic : UINT;
    stGlobPar  : ST_GlobPar;
    aMechPar   : ARRAY[1..GVL_Const.N_MECH] OF ST_MechPar;
    aValvePar  : ARRAY[1..GVL_Const.N_VALVE] OF ST_ValvePar;
    aBunkerPar : ARRAY[1..GVL_Const.N_BUNKER] OF ST_BunkerPar;
END_VAR

(* Бункер с датчиком верхнего уровня. Полный бункер ставит на паузу подающий участок
   маршрута; после освобождения и задержки uTRestart участок запускается снова. *)
FUNCTION_BLOCK FB_Bunker
VAR_INPUT
    xHasSF : BOOL;
    stIn   : ST_BunkerIn;
END_VAR
VAR_IN_OUT
    stHmi : ST_BunkerHmi;
    stPar : ST_BunkerPar;
END_VAR
VAR_OUTPUT
    xFull     : BOOL;
    xAlarm    : BOOL;
    xNewAlarm : BOOL;
END_VAR
VAR
    xDvu      : BOOL;
    wAct      : WORD;
    wAlm      : WORD;
    wSts      : WORD;
    uShDvu    : UINT;
    uShRst    : UINT;
    wShByp    : WORD;
    tonFull   : TON;
    tonClear  : TON;
END_VAR

            F_SyncUint(uMax := 600, uHmi := stHmi.uTDvu, uPar := stPar.uTDvu, uShadow := uShDvu);
F_SyncUint(uMax := GVL_Const.T_MAX_S, uHmi := stHmi.uTRestart, uPar := stPar.uTRestart, uShadow := uShRst);
F_SyncWord(wHmi := stHmi.wBypass, wPar := stPar.wBypass, wShadow := wShByp);

xDvu := stIn.xDVU AND (stPar.wBypass AND GVL_Const.BY_DVU) = 0;
tonFull(IN := xDvu, PT := F_Sec(stPar.uTDvu));
tonClear(IN := NOT xDvu, PT := F_Sec(stPar.uTRestart));
IF tonFull.Q THEN
    xFull := TRUE;
ELSIF tonClear.Q THEN
    xFull := FALSE;
END_IF

wAct := 0;
IF xHasSF AND NOT stIn.xSF THEN
    wAct := wAct OR GVL_Const.BA_SF;
END_IF
xNewAlarm := (wAct AND NOT wAlm) <> 0;
IF GVL.xReset THEN
    wAlm := wAct;
ELSE
    wAlm := wAlm OR wAct;
END_IF
xAlarm := wAlm <> 0;

wSts := 0;
IF stIn.xDVU THEN wSts := wSts OR GVL_Const.BS_DVU; END_IF
IF xFull THEN wSts := wSts OR GVL_Const.BS_FULL; END_IF
IF stIn.xDNU THEN wSts := wSts OR GVL_Const.BS_DNU; END_IF
IF (stPar.wBypass AND GVL_Const.BY_DVU) <> 0 THEN wSts := wSts OR GVL_Const.BS_BYPASS; END_IF
IF xAlarm THEN wSts := wSts OR GVL_Const.BS_ALARM; END_IF
stHmi.wSts := wSts;
stHmi.wAlm := wAlm;

          
END_FUNCTION_BLOCK

(* Механизм линии: двигатель прямого пуска, привод с ПЧ, заслонка с ПЧ или фотосепаратор.

   Режимы:
   - автомат (MODE_AUTO): работает по требованию маршрута. Пуск после задержки uTOn,
     когда все последующие механизмы уже работают (пуск от последнего к первому).
     Останов после задержки uTOff, когда нет требования и остановились все подающие
     механизмы (останов от первого к последнему);
   - ручной с панели (MODE_MAN): кнопки Пуск/Стоп, пуск разрешён только при работе
     последующих механизмов и неполных бункерах на выходе;
   - местный (MODE_LOCAL): ключ поста в "ручн.", кнопки поста;
   - наладка: ручной режим при GVL.xSetup - без блокировок и датчиков безопасности
     (кроме защит двигателя, аварийного стопа и аварии ПЧ).
   Переход между режимами безударный: команда работы сохраняется. *)
FUNCTION_BLOCK FB_Mech
VAR_INPUT
    stCfg       : ST_MechCfg;
    stIn        : ST_MechIn;
    xDemand     : BOOL;    (* требование активного маршрута *)
    xPredRun    : BOOL;    (* работает подающий механизм - удерживать в работе *)
    xSuccOkAuto : BOOL;    (* все последующие механизмы работают *)
    xSuccOkMan  : BOOL;    (* то же + бункеры на выходе не полны *)
    xPaused     : BOOL;    (* участок на паузе по ДВУ (для индикации) *)
END_VAR
VAR_IN_OUT
    stHmi : ST_MechHmi;
    stPar : ST_MechPar;
END_VAR
VAR_OUTPUT
    stOut     : ST_MechOut;
    xRun      : BOOL;      (* механизм в работе (для блокировок соседних) *)
    xCmd      : BOOL;      (* команда работы *)
    xReady    : BOOL;      (* готов к пуску в маршруте *)
    xAuto     : BOOL;
    xAlarm    : BOOL;
    xNewAlarm : BOOL;      (* появилась новая авария (один цикл) *)
END_VAR
VAR
    eMode      : INT;
    xManualReq : BOOL;
    xSetupNow  : BOOL;
    xStartReq  : BOOL;
    xStopReq   : BOOL;
    xMotorOn   : BOOL;     (* выход на двигатель был включен (предыдущий цикл) *)
    xSeqTrip   : BOOL;
    xSeqLatch  : BOOL;
    wAct       : WORD;
    wAlm       : WORD;
    xToDue     : BOOL;
    xOpened    : BOOL;
    xClosed    : BOOL;
    xGoOpen    : BOOL;
    xGoClose   : BOOL;
    xMoveBlock : BOOL;
    wSts       : WORD;
    uShTOn     : UINT;
    uShTOff    : UINT;
    uShTo      : UINT;
    wShByp     : WORD;
    tonStart   : TON;
    tonStop    : TON;
    tonDksRun  : TON;
    tonDksLost : TON;
    rtDks      : R_TRIG;
    tonDsl1    : TON;
    tonDsl2    : TON;
    tonDp      : TON;
    tonFb      : TON;
    tonMove    : TON;
    tpReset    : TP;
    rtCmd      : R_TRIG;
    ftCmd      : F_TRIG;
    tpOn       : TP;
    tpOff      : TP;
    rtLocStart : R_TRIG;
END_VAR

            (* ---- уставки панель <-> RETAIN ---- *)
F_SyncUint(uMax := GVL_Const.T_MAX_S, uHmi := stHmi.uTOn, uPar := stPar.uTOn, uShadow := uShTOn);
F_SyncUint(uMax := GVL_Const.T_MAX_S, uHmi := stHmi.uTOff, uPar := stPar.uTOff, uShadow := uShTOff);
F_SyncUint(uMax := 60000, uHmi := stHmi.uToInterval, uPar := stPar.uToInterval, uShadow := uShTo);
F_SyncWord(wHmi := stHmi.wBypass, wPar := stPar.wBypass, wShadow := wShByp);

(* ---- команды панели ---- *)
xStartReq := (stHmi.wCmd AND GVL_Const.C_START) <> 0;
xStopReq := (stHmi.wCmd AND GVL_Const.C_STOP) <> 0;
IF (stHmi.wCmd AND GVL_Const.C_RESET_TO) <> 0 THEN
    stPar.udSecSinceTO := 0;
END_IF
stHmi.wCmd := stHmi.wCmd AND NOT (GVL_Const.C_START OR GVL_Const.C_STOP OR GVL_Const.C_RESET_TO);

(* механизм, занятый маршрутом, в ручной режим с панели не переводится *)
IF xDemand THEN
    stHmi.wCmd := stHmi.wCmd AND NOT GVL_Const.C_MANUAL;
END_IF
xManualReq := (stHmi.wCmd AND GVL_Const.C_MANUAL) <> 0;

IF stCfg.xHasLocal AND stIn.xLocal THEN
    eMode := GVL_Const.MODE_LOCAL;
ELSIF xManualReq THEN
    eMode := GVL_Const.MODE_MAN;
ELSE
    eMode := GVL_Const.MODE_AUTO;
END_IF
xSetupNow := GVL.xSetup AND eMode = GVL_Const.MODE_MAN;
xAuto := eMode = GVL_Const.MODE_AUTO;

(* ---- аварии ---- *)
wAct := 0;
IF stCfg.xHasQF AND NOT stIn.xQF THEN
    wAct := wAct OR GVL_Const.A_QF;
END_IF

tonDksRun(IN := xMotorOn AND stCfg.eDks <> GVL_Const.DKS_NONE, PT := F_Sec(GVL_Retain.stGlobPar.uTDksGrace));
rtDks(CLK := stIn.xDKS);
IF stCfg.eDks = GVL_Const.DKS_PULSE THEN
    (* таймер перезапускается каждым фронтом импульса *)
    tonDksLost(IN := tonDksRun.Q AND NOT rtDks.Q,
               PT := UDINT_TO_TIME(UINT_TO_UDINT(GVL_Retain.stGlobPar.uTDksPulse) * 100));
ELSE
    tonDksLost(IN := tonDksRun.Q AND NOT stIn.xDKS,
               PT := UDINT_TO_TIME(UINT_TO_UDINT(GVL_Retain.stGlobPar.uTDksPulse) * 100));
END_IF
IF tonDksLost.Q AND (stPar.wBypass AND GVL_Const.BY_DKS) = 0 THEN
    wAct := wAct OR GVL_Const.A_DKS;
END_IF

(* сбег ленты контролируется и на стоящей нории: пуск со сбежавшей лентой запрещён *)
tonDsl1(IN := stCfg.xHasDSL AND NOT stIn.xDSL1, PT := T#1S);
IF tonDsl1.Q AND (stPar.wBypass AND GVL_Const.BY_DSL1) = 0 THEN
    wAct := wAct OR GVL_Const.A_DSL1;
END_IF
tonDsl2(IN := stCfg.xHasDSL AND NOT stIn.xDSL2, PT := T#1S);
IF tonDsl2.Q AND (stPar.wBypass AND GVL_Const.BY_DSL2) = 0 THEN
    wAct := wAct OR GVL_Const.A_DSL2;
END_IF
tonDp(IN := stCfg.xHasDP AND NOT stIn.xDP, PT := T#2S);
IF tonDp.Q AND (stPar.wBypass AND GVL_Const.BY_DP) = 0 THEN
    wAct := wAct OR GVL_Const.A_DP;
END_IF

IF stCfg.xHasEStop AND NOT stIn.xEStop THEN
    wAct := wAct OR GVL_Const.A_ESTOP;
END_IF
(* местный "Стоп" при работе от панели/маршрута: механизм уже отключен аппаратно *)
IF stCfg.xHasLocal AND NOT stIn.xLocStop AND eMode <> GVL_Const.MODE_LOCAL AND (xCmd OR xDemand) THEN
    wAct := wAct OR GVL_Const.A_LOCSTOP;
END_IF

CASE stCfg.eKind OF
GVL_Const.K_FC:
    IF stIn.xFcFault THEN
        wAct := wAct OR GVL_Const.A_FC;
    END_IF
    tonFb(IN := xMotorOn AND NOT stIn.xFcReady, PT := F_Sec(GVL_Retain.stGlobPar.uTFcFb));
    IF tonFb.Q THEN
        wAct := wAct OR GVL_Const.A_FCFB;
    END_IF
GVL_Const.K_GATE:
    IF stIn.xFcFault THEN
        wAct := wAct OR GVL_Const.A_FC;
    END_IF
    tonMove(IN := stOut.qOpen OR stOut.qClose, PT := F_Sec(GVL_Retain.stGlobPar.uTGateMove));
    IF tonMove.Q THEN
        wAct := wAct OR GVL_Const.A_MOVE;
    END_IF
    IF stIn.xFb1 AND stIn.xFb2 THEN
        wAct := wAct OR GVL_Const.A_POS;
    END_IF
GVL_Const.K_FS:
    IF stIn.xErr THEN
        wAct := wAct OR GVL_Const.A_FSERR;
    END_IF
    tonFb(IN := xCmd AND NOT stIn.xFb1, PT := F_Sec(GVL_Retain.stGlobPar.uTFsStart));
    IF tonFb.Q THEN
        wAct := wAct OR GVL_Const.A_FSFB;
    END_IF
END_CASE

IF xSetupNow THEN
    wAct := wAct AND GVL_Const.A_HARD;
END_IF

(* фиксация аварий до сброса *)
xNewAlarm := (wAct AND NOT wAlm) <> 0;
IF GVL.xReset THEN
    wAlm := wAct;
    xSeqLatch := FALSE;
ELSE
    wAlm := wAlm OR wAct;
END_IF
xAlarm := wAlm <> 0;

(* ---- готовность к работе в маршруте ---- *)
xReady := NOT xAlarm AND xAuto AND GVL.xGlobalOk
    AND (NOT stCfg.xHasLocal OR stIn.xLocStop)
    AND (NOT stCfg.xHasEStop OR stIn.xEStop)
    AND (stCfg.eKind <> GVL_Const.K_FS
         OR (stIn.xFb2 AND (stIn.xAux OR (stPar.wBypass AND GVL_Const.BY_AUX) <> 0)));

(* ---- команда работы ---- *)
rtLocStart(CLK := stIn.xLocStart);
CASE eMode OF
GVL_Const.MODE_AUTO:
    tonStart(IN := xDemand AND xSuccOkAuto AND xReady AND NOT xCmd, PT := F_Sec(stPar.uTOn));
    IF tonStart.Q THEN
        xCmd := TRUE;
        xSeqLatch := FALSE;
    END_IF
    tonStop(IN := xCmd AND NOT xDemand AND NOT xPredRun, PT := F_Sec(stPar.uTOff));
    IF tonStop.Q THEN
        xCmd := FALSE;
    END_IF
    xSeqTrip := NOT xSuccOkAuto;

GVL_Const.MODE_MAN:
    tonStart(IN := FALSE);
    tonStop(IN := FALSE);
    IF xStartReq AND NOT xAlarm AND GVL.xGlobalOk AND (xSuccOkMan OR xSetupNow) THEN
        xCmd := TRUE;
        xSeqLatch := FALSE;
    END_IF
    IF xStopReq THEN
        xCmd := FALSE;
    END_IF
    xSeqTrip := NOT xSuccOkMan AND NOT xSetupNow;

GVL_Const.MODE_LOCAL:
    tonStart(IN := FALSE);
    tonStop(IN := FALSE);
    IF rtLocStart.Q AND NOT xAlarm AND stIn.xLocStop THEN
        xCmd := TRUE;
    END_IF
    IF NOT stIn.xLocStop THEN
        xCmd := FALSE;
    END_IF
    xSeqTrip := FALSE;
END_CASE

(* заслонка управляется в местном и ручном режимах кнопками открыть/закрыть, см. ниже *)
IF stCfg.eKind = GVL_Const.K_GATE AND eMode <> GVL_Const.MODE_AUTO THEN
    xCmd := FALSE;
    xSeqTrip := FALSE;
END_IF

IF xCmd AND xSeqTrip THEN
    xSeqLatch := TRUE;
END_IF
(* аварийный стоп, пожар, фазы, отключение цепи управления - останов сразу, без задержек *)
IF xAlarm OR NOT GVL.xGlobalOk OR xSeqTrip THEN
    xCmd := FALSE;
END_IF

(* ---- исполнительная часть ---- *)
stOut.qRun := FALSE;
stOut.qPower := FALSE;
stOut.qOpen := FALSE;
stOut.qClose := FALSE;
stOut.qEnable := FALSE;
tpReset(IN := GVL.xReset, PT := T#1S);
stOut.qReset := tpReset.Q;
rtCmd(CLK := xCmd);
ftCmd(CLK := xCmd);
tpOn(IN := rtCmd.Q AND stCfg.eKind = GVL_Const.K_FS, PT := T#1S);
tpOff(IN := ftCmd.Q AND stCfg.eKind = GVL_Const.K_FS, PT := T#1S);
stOut.qOn := tpOn.Q;
stOut.qOff := tpOff.Q;
xOpened := stIn.xFb1 AND NOT stIn.xFb2;
xClosed := stIn.xFb2 AND NOT stIn.xFb1;

CASE stCfg.eKind OF
GVL_Const.K_DOL:
    stOut.qRun := xCmd;
    xRun := xCmd;
    xMotorOn := xCmd;

GVL_Const.K_FC:
    stOut.qPower := GVL.xSysOn AND (NOT stCfg.xHasQF OR stIn.xQF);
    stOut.qRun := xCmd AND stOut.qPower;
    xRun := stOut.qRun;
    xMotorOn := stOut.qRun;

GVL_Const.K_GATE:
    stOut.qPower := GVL.xSysOn AND (NOT stCfg.xHasQF OR stIn.xQF);
    CASE eMode OF
    GVL_Const.MODE_AUTO:
        xGoOpen := xCmd;
        xGoClose := NOT xCmd;
    GVL_Const.MODE_MAN:
        xGoOpen := (stHmi.wCmd AND GVL_Const.C_OPEN) <> 0 AND (xSuccOkMan OR xSetupNow);
        xGoClose := (stHmi.wCmd AND GVL_Const.C_CLOSE) <> 0;
    ELSE
        xGoOpen := stIn.xLocOpen AND stIn.xLocStop;
        xGoClose := stIn.xLocClose AND stIn.xLocStop;
    END_CASE
    (* при общей аварии заслонка только закрывается - прекращение подачи продукта *)
    xGoOpen := xGoOpen AND GVL.xGlobalOk;
    (* ход прекращается при аварии привода или концевиков до сброса *)
    xMoveBlock := (wAlm AND (GVL_Const.A_QF OR GVL_Const.A_FC OR GVL_Const.A_MOVE OR GVL_Const.A_POS)) <> 0
        OR NOT stOut.qPower;
    stOut.qOpen := xGoOpen AND NOT xGoClose AND NOT xOpened AND NOT xMoveBlock;
    stOut.qClose := xGoClose AND NOT xGoOpen AND NOT xClosed AND NOT xMoveBlock;
    (* проём не закрыт - продукт может поступать на норию *)
    xRun := stOut.qOpen OR xOpened OR (NOT xClosed AND NOT xAlarm);
    xMotorOn := stOut.qOpen OR stOut.qClose;

GVL_Const.K_FS:
    stOut.qEnable := xCmd AND stIn.xFb1;
    xRun := xCmd AND stIn.xFb1;
    xMotorOn := xRun;
END_CASE

(* ---- моточасы ---- *)
IF xMotorOn AND GVL.xPulse1s THEN
    stPar.udSecTotal := stPar.udSecTotal + 1;
    stPar.udSecSinceTO := stPar.udSecSinceTO + 1;
END_IF
stHmi.uHoursTotal := UDINT_TO_UINT(MIN(stPar.udSecTotal / 3600, 65535));
stHmi.uMinutes := UDINT_TO_UINT((stPar.udSecTotal / 60) MOD 60);
stHmi.uHoursSinceTO := UDINT_TO_UINT(MIN(stPar.udSecSinceTO / 3600, 65535));
xToDue := stPar.uToInterval > 0 AND stPar.udSecSinceTO / 3600 >= UINT_TO_UDINT(stPar.uToInterval);

(* ---- состояние для панели ---- *)
wSts := 0;
IF xRun THEN wSts := wSts OR GVL_Const.S_RUN; END_IF
IF xCmd THEN wSts := wSts OR GVL_Const.S_CMD; END_IF
IF xReady THEN wSts := wSts OR GVL_Const.S_READY; END_IF
IF xAlarm THEN wSts := wSts OR GVL_Const.S_ALARM; END_IF
IF eMode = GVL_Const.MODE_LOCAL THEN wSts := wSts OR GVL_Const.S_LOCAL; END_IF
IF eMode = GVL_Const.MODE_MAN THEN wSts := wSts OR GVL_Const.S_MANUAL; END_IF
IF xSetupNow THEN wSts := wSts OR GVL_Const.S_SETUP; END_IF
IF tonStart.IN AND NOT xCmd THEN wSts := wSts OR GVL_Const.S_STARTING; END_IF
IF tonStop.IN THEN wSts := wSts OR GVL_Const.S_STOPPING; END_IF
IF xDemand THEN wSts := wSts OR GVL_Const.S_DEMAND; END_IF
IF xPaused THEN wSts := wSts OR GVL_Const.S_PAUSE; END_IF
IF xToDue THEN wSts := wSts OR GVL_Const.S_TO_DUE; END_IF
IF xOpened THEN wSts := wSts OR GVL_Const.S_OPENED; END_IF
IF xClosed THEN wSts := wSts OR GVL_Const.S_CLOSED; END_IF
IF xSeqLatch THEN wSts := wSts OR GVL_Const.S_SEQ_TRIP; END_IF
IF xSuccOkMan THEN wSts := wSts OR GVL_Const.S_SUCC_OK; END_IF
stHmi.wSts := wSts;
stHmi.wAlm := wAlm;

IF xAlarm THEN
    stHmi.iState := 4;
ELSIF eMode = GVL_Const.MODE_LOCAL THEN
    stHmi.iState := 5;
ELSIF tonStop.IN THEN
    stHmi.iState := 3;
ELSIF xRun THEN
    stHmi.iState := 2;
ELSIF tonStart.IN THEN
    stHmi.iState := 1;
ELSE
    stHmi.iState := 0;
END_IF

          
END_FUNCTION_BLOCK

(* Переключатель потока ППМ-2 с электроприводом (поз.12(1)..12(4)) и
   механизм промежуточной выгрузки Z-нории поз.26 (пневмораспределитель 49YA1/49YA2).
   Выход держится до срабатывания датчика положения. Положение задаёт маршрут;
   в ручном режиме - кнопки панели, если подающий механизм стоит. *)
FUNCTION_BLOCK FB_Valve
VAR_INPUT
    xHasSF  : BOOL;
    stIn    : ST_ValveIn;
    iTarget : INT;      (* 0 - нет задания маршрута, 1/2 - положение *)
    xFlow   : BOOL;     (* подающий механизм работает *)
END_VAR
VAR_IN_OUT
    stHmi : ST_ValveHmi;
    stPar : ST_ValvePar;
END_VAR
VAR_OUTPUT
    stOut     : ST_ValveOut;
    iPos      : INT;    (* 0 - не определено, 1, 2 *)
    xReady    : BOOL;
    xAlarm    : BOOL;
    xNewAlarm : BOOL;
END_VAR
VAR
    iGoal    : INT;
    xManual  : BOOL;
    xReq1    : BOOL;
    xReq2    : BOOL;
    xMove1   : BOOL;
    xMove2   : BOOL;
    wAct     : WORD;
    wAlm     : WORD;
    wSts     : WORD;
    uShMove  : UINT;
    tonMove  : TON;
    tofQ1    : TOF;
    tofQ2    : TOF;
END_VAR

            F_SyncUint(uMax := 600, uHmi := stHmi.uTMove, uPar := stPar.uTMove, uShadow := uShMove);

IF stIn.xS1 AND NOT stIn.xS2 THEN
    iPos := 1;
ELSIF stIn.xS2 AND NOT stIn.xS1 THEN
    iPos := 2;
ELSE
    iPos := 0;
END_IF

(* ---- аварии ---- *)
wAct := 0;
IF xHasSF AND NOT stIn.xSF THEN
    wAct := wAct OR GVL_Const.VA_SF;
END_IF
tonMove(IN := stOut.q1 OR stOut.q2, PT := F_Sec(stPar.uTMove));
IF tonMove.Q THEN
    wAct := wAct OR GVL_Const.VA_TIMEOUT;
END_IF
IF stIn.xS1 AND stIn.xS2 THEN
    wAct := wAct OR GVL_Const.VA_BOTH;
END_IF
xNewAlarm := (wAct AND NOT wAlm) <> 0;
IF GVL.xReset THEN
    wAlm := wAct;
ELSE
    wAlm := wAlm OR wAct;
END_IF
xAlarm := wAlm <> 0;

(* ---- задание положения ---- *)
IF iTarget <> 0 THEN
    stHmi.wCmd := stHmi.wCmd AND NOT GVL_Const.VC_MANUAL;
END_IF
xManual := (stHmi.wCmd AND GVL_Const.VC_MANUAL) <> 0;
xReq1 := (stHmi.wCmd AND GVL_Const.VC_POS1) <> 0;
xReq2 := (stHmi.wCmd AND GVL_Const.VC_POS2) <> 0;
stHmi.wCmd := stHmi.wCmd AND NOT (GVL_Const.VC_POS1 OR GVL_Const.VC_POS2);

IF iTarget <> 0 THEN
    iGoal := iTarget;
ELSIF xManual THEN
    IF NOT xFlow OR GVL.xSetup THEN
        IF xReq1 THEN
            iGoal := 1;
        ELSIF xReq2 THEN
            iGoal := 2;
        END_IF
    END_IF
ELSE
    iGoal := 0;
END_IF

xMove1 := iGoal = 1 AND iPos <> 1 AND NOT xAlarm AND GVL.xGlobalOk;
xMove2 := iGoal = 2 AND iPos <> 2 AND NOT xAlarm AND GVL.xGlobalOk;
(* пауза 0,5 с при реверсе привода *)
stOut.q1 := xMove1 AND NOT tofQ2.Q;
stOut.q2 := xMove2 AND NOT tofQ1.Q AND NOT stOut.q1;
tofQ1(IN := stOut.q1, PT := T#500MS);
tofQ2(IN := stOut.q2, PT := T#500MS);

xReady := NOT xAlarm AND NOT xManual;

wSts := 0;
IF iPos = 1 THEN wSts := wSts OR GVL_Const.VS_POS1; END_IF
IF iPos = 2 THEN wSts := wSts OR GVL_Const.VS_POS2; END_IF
IF stOut.q1 OR stOut.q2 THEN wSts := wSts OR GVL_Const.VS_MOVING; END_IF
IF xAlarm THEN wSts := wSts OR GVL_Const.VS_ALARM; END_IF
IF xManual THEN wSts := wSts OR GVL_Const.VS_MANUAL; END_IF
IF iTarget <> 0 THEN wSts := wSts OR GVL_Const.VS_ROUTE; END_IF
IF xFlow THEN wSts := wSts OR GVL_Const.VS_FLOW; END_IF
stHmi.wSts := wSts;
stHmi.wAlm := wAlm;

          
END_FUNCTION_BLOCK

(* Связи "кто на кого подаёт" при заданных положениях клапанов.
   Используется для блокировок (с фактическими положениями) и для определения состава
   маршрутов (с положениями из ROUTE_VALVE). Возвращает число связей. *)
FUNCTION F_BuildLinks : INT
VAR_IN_OUT
    aPos   : ARRAY[1..GVL_Const.N_VALVE] OF INT;
    aLinks : ARRAY[1..GVL_Const.N_LINK] OF ST_Link;
END_VAR
VAR
    n : INT;
END_VAR
VAR CONSTANT
    M : INT := 0;   (* LT_MECH *)
    B : INT := 1;   (* LT_BUNKER *)
    X : INT := 2;   (* LT_INVALID *)
END_VAR

            (* ---- приёмное отделение и МУЗ ---- *)
n := n + 1; aLinks[n] := F_Link(GVL_Const.M_GATE1, M, GVL_Const.M_N3, TRUE);
n := n + 1; aLinks[n] := F_Link(GVL_Const.M_N3, B, GVL_Const.B_B4, TRUE);
n := n + 1; aLinks[n] := F_Link(GVL_Const.M_MUZ5_FD, M, GVL_Const.M_MUZ5, TRUE);
n := n + 1; aLinks[n] := F_Link(GVL_Const.M_MUZ5, M, GVL_Const.M_N7, TRUE);
n := n + 1; aLinks[n] := F_Link(GVL_Const.M_MUZ5, M, GVL_Const.M_SH32, FALSE);    (* неиспользуемые отходы 32-31-30 *)
n := n + 1; aLinks[n] := F_Link(GVL_Const.M_MUZ5, M, GVL_Const.M_KC35, FALSE);    (* используемые отходы 35-34 *)
n := n + 1; aLinks[n] := F_Link(GVL_Const.M_MUZ5, M, GVL_Const.M_FAN6, FALSE);
n := n + 1; aLinks[n] := F_Link(GVL_Const.M_FAN6, M, GVL_Const.M_SL6, FALSE);
n := n + 1; aLinks[n] := F_Link(GVL_Const.M_N7, B, GVL_Const.B_B8, TRUE);

(* ---- ТОР-18 ---- *)
n := n + 1; aLinks[n] := F_Link(GVL_Const.M_TOR9_FD, M, GVL_Const.M_TOR9, TRUE);
n := n + 1; aLinks[n] := F_Link(GVL_Const.M_TOR9, M, GVL_Const.M_N11, TRUE);
n := n + 1; aLinks[n] := F_Link(GVL_Const.M_TOR9, M, GVL_Const.M_SH31, FALSE);    (* неиспользуемые 31-30 *)
n := n + 1; aLinks[n] := F_Link(GVL_Const.M_TOR9, M, GVL_Const.M_KC35, FALSE);
n := n + 1; aLinks[n] := F_Link(GVL_Const.M_TOR9, M, GVL_Const.M_FAN10, FALSE);
n := n + 1; aLinks[n] := F_Link(GVL_Const.M_FAN10, M, GVL_Const.M_SL10, FALSE);

(* нория 11 -> 12(1) -> TORBA 13(1) | 12(2) -> БТ | растариватель 15(1) -> нория 16 *)
CASE aPos[GVL_Const.V_V12_1] OF
1:
    n := n + 1; aLinks[n] := F_Link(GVL_Const.M_N11, B, GVL_Const.B_T13_1, TRUE);
2:
    CASE aPos[GVL_Const.V_V12_2] OF
    1:
        n := n + 1; aLinks[n] := F_Link(GVL_Const.M_N11, M, GVL_Const.M_BT14_1, TRUE);
        n := n + 1; aLinks[n] := F_Link(GVL_Const.M_N11, M, GVL_Const.M_BT14_2, TRUE);
    2:
        n := n + 1; aLinks[n] := F_Link(GVL_Const.M_N11, M, GVL_Const.M_N16, TRUE);
    ELSE
        n := n + 1; aLinks[n] := F_Link(GVL_Const.M_N11, X, 0, TRUE);
    END_CASE
ELSE
    n := n + 1; aLinks[n] := F_Link(GVL_Const.M_N11, X, 0, TRUE);
END_CASE

(* ---- блок триерный ---- *)
n := n + 1; aLinks[n] := F_Link(GVL_Const.M_BT14_1, M, GVL_Const.M_N16, TRUE);
n := n + 1; aLinks[n] := F_Link(GVL_Const.M_BT14_2, M, GVL_Const.M_N16, TRUE);
n := n + 1; aLinks[n] := F_Link(GVL_Const.M_BT14_1, M, GVL_Const.M_KC36, FALSE);  (* отходы 36-35-34 *)
n := n + 1; aLinks[n] := F_Link(GVL_Const.M_BT14_2, M, GVL_Const.M_KC36, FALSE);

(* нория 16 -> 12(3) -> бункер 17 (КСП) | нория 20 *)
CASE aPos[GVL_Const.V_V12_3] OF
1:
    n := n + 1; aLinks[n] := F_Link(GVL_Const.M_N16, B, GVL_Const.B_B17, TRUE);
2:
    n := n + 1; aLinks[n] := F_Link(GVL_Const.M_N16, M, GVL_Const.M_N20, TRUE);
ELSE
    n := n + 1; aLinks[n] := F_Link(GVL_Const.M_N16, X, 0, TRUE);
END_CASE

(* ---- КСП-11М ---- *)
n := n + 1; aLinks[n] := F_Link(GVL_Const.M_KSP18_FD, M, GVL_Const.M_KSP18, TRUE);
n := n + 1; aLinks[n] := F_Link(GVL_Const.M_KSP18, M, GVL_Const.M_N20, TRUE);
n := n + 1; aLinks[n] := F_Link(GVL_Const.M_KSP18, M, GVL_Const.M_SH33, FALSE);   (* неиспользуемые 33-31-30 *)
n := n + 1; aLinks[n] := F_Link(GVL_Const.M_KSP18, M, GVL_Const.M_KC35, FALSE);
n := n + 1; aLinks[n] := F_Link(GVL_Const.M_KSP18, M, GVL_Const.M_FAN19, FALSE);
n := n + 1; aLinks[n] := F_Link(GVL_Const.M_FAN19, M, GVL_Const.M_SL19, FALSE);
n := n + 1; aLinks[n] := F_Link(GVL_Const.M_N20, B, GVL_Const.B_B22, TRUE);

(* нория 21 -> 12(4) -> бункер 22 (СП) | Z-нория 26 *)
CASE aPos[GVL_Const.V_V12_4] OF
1:
    n := n + 1; aLinks[n] := F_Link(GVL_Const.M_N21, B, GVL_Const.B_B22, TRUE);
2:
    n := n + 1; aLinks[n] := F_Link(GVL_Const.M_N21, M, GVL_Const.M_ZN26, TRUE);
ELSE
    n := n + 1; aLinks[n] := F_Link(GVL_Const.M_N21, X, 0, TRUE);
END_CASE

(* ---- СП-200 ---- *)
n := n + 1; aLinks[n] := F_Link(GVL_Const.M_SP24_DRV, M, GVL_Const.M_ZN26, TRUE);
n := n + 1; aLinks[n] := F_Link(GVL_Const.M_SP24_DRV, M, GVL_Const.M_KC36, FALSE);
n := n + 1; aLinks[n] := F_Link(GVL_Const.M_SP24_DRV, M, GVL_Const.M_SP24_FAN, FALSE);
n := n + 1; aLinks[n] := F_Link(GVL_Const.M_SP24_FAN, M, GVL_Const.M_FAN25, FALSE);
n := n + 1; aLinks[n] := F_Link(GVL_Const.M_FAN25, M, GVL_Const.M_SL25, FALSE);

(* Z-нория 26 -> выгрузка включена: TORBA 13(2) | выключена: бункер фотосепаратора *)
CASE aPos[GVL_Const.V_V49] OF
1:
    n := n + 1; aLinks[n] := F_Link(GVL_Const.M_ZN26, B, GVL_Const.B_T13_2, TRUE);
2:
    n := n + 1; aLinks[n] := F_Link(GVL_Const.M_ZN26, B, GVL_Const.B_B27, TRUE);
ELSE
    n := n + 1; aLinks[n] := F_Link(GVL_Const.M_ZN26, X, 0, TRUE);
END_CASE

(* ---- фотосепаратор (отходы - напрямую в рамку Биг-Бег) ---- *)
n := n + 1; aLinks[n] := F_Link(GVL_Const.M_FS27, M, GVL_Const.M_ZN29, TRUE);
n := n + 1; aLinks[n] := F_Link(GVL_Const.M_FS27, M, GVL_Const.M_FAN28, FALSE);
n := n + 1; aLinks[n] := F_Link(GVL_Const.M_FAN28, M, GVL_Const.M_SL28, FALSE);
n := n + 1; aLinks[n] := F_Link(GVL_Const.M_ZN29, B, GVL_Const.B_T13_2, TRUE);

(* ---- конвейеры отходов ---- *)
n := n + 1; aLinks[n] := F_Link(GVL_Const.M_SH32, M, GVL_Const.M_SH31, FALSE);
n := n + 1; aLinks[n] := F_Link(GVL_Const.M_SH33, M, GVL_Const.M_SH31, FALSE);
n := n + 1; aLinks[n] := F_Link(GVL_Const.M_SH31, M, GVL_Const.M_SH30, FALSE);
n := n + 1; aLinks[n] := F_Link(GVL_Const.M_KC36, M, GVL_Const.M_KC35, FALSE);
n := n + 1; aLinks[n] := F_Link(GVL_Const.M_KC35, M, GVL_Const.M_KC34, FALSE);

F_BuildLinks := n;

          
END_FUNCTION

FUNCTION F_Link : ST_Link
VAR_INPUT
    iFrom    : INT;
    eTo      : INT;
    iTo      : INT;
    xProduct : BOOL;
END_VAR

            F_Link.iFrom := iFrom;
F_Link.eTo := eTo;
F_Link.iTo := iTo;
F_Link.xProduct := xProduct;

          
END_FUNCTION

(* Секунды (UINT) -> TIME *)
FUNCTION F_Sec : TIME
VAR_INPUT
    uSec : UINT;
END_VAR

            F_Sec := UDINT_TO_TIME(UINT_TO_UDINT(uSec) * 1000);

          
END_FUNCTION

(* Уставка в RETAIN <-> регистр панели.
   Если панель изменила регистр (он отличается от последнего выданного значения) -
   принять новое значение с ограничением, затем выдать уставку обратно в регистр. *)
FUNCTION F_SyncUint : BOOL
VAR_INPUT
    uMax : UINT;
END_VAR
VAR_IN_OUT
    uHmi    : UINT;
    uPar    : UINT;
    uShadow : UINT;
END_VAR

            IF uHmi <> uShadow THEN
    uPar := MIN(uHmi, uMax);
    F_SyncUint := TRUE;
END_IF
uHmi := uPar;
uShadow := uPar;

          
END_FUNCTION

FUNCTION F_SyncWord : BOOL
VAR_IN_OUT
    wHmi    : WORD;
    wPar    : WORD;
    wShadow : WORD;
END_VAR

            IF wHmi <> wShadow THEN
    wPar := wHmi;
    F_SyncWord := TRUE;
END_IF
wHmi := wPar;
wShadow := wPar;

          
END_FUNCTION

(* Главная программа. Вызывается из задачи MAST (циклическая, 20 мс). *)
PROGRAM PLC_PRG

            PRG_Inputs();
PRG_System();
PRG_Topology();
PRG_Routes();
PRG_Mechs();
PRG_Outputs();

          
END_PROGRAM

(* Сгенерировано gen/gen_io.py. Физические входы -> логические сигналы.
   Полярность датчиков - константы CFG_* в GVL_Const. *)
PROGRAM PRG_Inputs

